(* IEC 61131-3 sources: daoli-st-library/DL_MathData (part 30) *)

(* ---- FB_DL_StringTokenStream.st ---- *)
(*==============================================================================
 * 组件名称 (Component)  : FB_DL_StringTokenStream
 * 所属子库 (Sublibrary) : DL_MathData
 * 当前版本 (Version)    : 1.0.1
 * 兼容性   (Platform)   : CODESYS 3.5 / TwinCAT 3 / 汇川 InoProShop / Machine Expert
 *                         仅依赖 Standard.library（LEN / FIND / LEFT / MID / R_TRIG）
 * 功能描述 (Function)   : 按 1~4 字符分隔符把一条定长报文逐段取出，每次触发输出一段，
 *                         跨扫描周期推进。用于扫码枪、称重仪表、在线分析仪这类
 *                         「字段长度不固定、帧总长有限」的报文解析。
 *                         本件最重要的语义：**连续分隔符产生空段，空段仍占一个序号**，
 *                         绝不跳过、绝不合并 —— 现场手写取段程序最典型的故障就是空字段
 *                         被吞掉导致后续字段整体错位（第 3 段显示成第 4 段的值）。
 *                         流式推进的另一目的是把「一次解析整帧」的耗时摊到多拍，
 *                         不让长报文的串操作撑爆扫描周期。
 * 出口契约 (Exit)       : sToken / nTokenIdx / bValidToken 为「本拍产出」，bDone 表示帧已读完
 *                          （读完后保持 TRUE，直到重装载或复位）。故障级锁存只由 021C /
 *                         021D / 021E 三码置位，bReset 上升沿统一清故障并回空闲。
 *                         调用约定：bNext 上升沿后**下一拍**产出该段（状态机一相一拍，
 *                         便于上层在「请求」与「结果」之间插入握手超时判断）。
 * 开源溯源 (Origin)     : 来源标签 lgf-datahandling。许可证：LGF 为免费闭源发布，未取得源码，
 *                         不构成衍生作品。借鉴点仅为字符串族「定长缓冲 + 原地操作、
 *                         不做动态分配」的参数域契约。
 *                         clean-room 独立实现：流式状态机、空段语义、段数上限策略、
 *                         帧改写判据、错误码全部自有——该类库并无流式分词器可参考。
 * 码位说明 (Codes)      : 信息级 16#0001_013A（空段）/ 013B（段长超限已截断）/ 013C（末段后
 *                         再取）；故障级 16#0001_021C（分隔符为空）/ 021D（段数超上限）/
 *                         021E（非法相位兜底）。共 6 码，全部落在 R12 计划第 1.2 节本件码段内。
 * 依赖     (Depends)    : 无 DL_ 内部依赖；Standard.library: LEN / FIND / LEFT / MID / R_TRIG
 * 红线自检 (Redline)    : 1 ✓ 零全局变量表依赖、零外部变量声明、零物理地址
 *                         2 ✓ 纯 IEC 61131-3，无指针、无厂商库、无动态内存
 *                         3 ✓ 分隔符空硬闸、段数上限锁故障、段长截断、游标全程夹在帧内
 *                         4 ✓ 全变量中英双语同行注释
 *                         5 ✓ 四态 ENUM + CASE 全覆盖 + ELSE 兜底（021E）
 *                         6 ✓ R_TRIG 实例在 CASE 之外每拍无条件刷新
 *                         7 ✓ END_FUNCTION_BLOCK 位于文件最后有效行
 * 规格偏离留档 (Deviation):
 *   D1 计划 3.7 节内部变量表列有 fbTrigFrame（帧变化沿实例）。实测「等长改写」场景下
 *      帧变化必须逐字符比较才能判出，边沿实例反而会漏判（连续两拍都不同则不再产生上升沿），
 *      故本实现只保留 fbTrigNext / fbTrigReset 两个实例，帧变化判据改为逐字符比较，
 *      不设 fbTrigFrame，避免出现「声明了却不参与判决」的死变量。
 *   D2 计划写「bDone 单拍脉冲」，同节边界条款又写「bDone 保持 TRUE」。本实现取后者
 *      （保持到重装载或复位），理由：上层若每拍轮询 bDone，单拍脉冲极易漏采。
 * 修订历史 (Revision)   :
 *   2026-11-15  v1.0.0  首版入库（R12 · Level 0/1 DL_MathData 字符串族）
 *   2026-11-15  v1.0.1  终审定点修复 A-D02：取段相位（eDraining）入口用锁存帧长度
 *      重算 nFrameLen，与全局帧长度判据（段 3 跟随实时入参）解耦。原实现取段时用
 *      实时帧长度做边界与 MID 长度，却对锁存副本切片，调用方中途改写帧即可能产出
 *      「有效但为空」的假段（nSegLen 取自实时帧、字符取自短一截的锁存帧）
 *============================================================================*)

(*-----------------------------------------------------------------------------
 * 枚举: E_DL_TokenPhase（归属 DL_MathData，与本功能块同文件）
 * 含义: 分词流式解析的离散相位。步长留空位，便于后续插态而不破坏既有工程数值。
 *----------------------------------------------------------------------------*)
TYPE E_DL_TokenPhase :
(
    eIdle     := 0,    // 空闲：等待使能与分隔符校验 / Idle: waiting for enable and delimiter check
    eReady    := 10,   // 就绪：等待帧装载或下一次取段请求 / Ready: waiting for frame load or next request
    eDraining := 20,   // 取段：本拍切出一段并推进游标 / Draining: cut one segment and advance the cursor
    eFault    := 99    // 故障：分隔符为空或段数超限，输出冻结 / Fault: bad delimiter or token overflow
);
END_TYPE

(*==============================================================================
 * 功能块: FB_DL_StringTokenStream
 * 调用约定: 每个扫描周期无条件调用一次；bEnable 为 FALSE 时内部相位与全部出口冻结。
 * 无状态泄漏: 全部状态驻留于实例私有 VAR，零全局引用，可多实例并行解析多条报文。
 *============================================================================*)
FUNCTION_BLOCK FB_DL_StringTokenStream
VAR_INPUT
    bEnable       : BOOL;                        // 使能，FALSE 时冻结游标并保持全部输出 / Enable, freezes the cursor when FALSE
    bReset        : BOOL;                        // 上升沿复位到帧起点并清故障 / Rising edge rewinds to the frame start
    sFrame        : STRING(255);                 // 待分词报文，内容变化自动重装载 / Frame to tokenise, reloaded on change
    sDelimiter    : STRING(4);                   // 分隔符（1~4 字符），空 = 故障 / Delimiter of one to four characters
    bNext         : BOOL;                        // 上升沿取下一段 / Rising edge advances to the next token
    nMaxTokenLen  : INT := 32;                   // 单段最大长度 [字符]，域 1~64 / Maximum token length, 1..64
    nMaxTokens    : INT := 32;                   // 单帧最大段数 [段]，域 1~64 / Maximum token count, 1..64
END_VAR
VAR_OUTPUT
    sToken        : STRING(64);                  // 本段内容，超长截断 / Current token, truncated when too long
    nTokenIdx     : INT;                         // 本段序号，1 起 [索引] / Token index, one based
    nTokenCount   : INT;                         // 本帧已产出段数 [段] / Tokens produced so far
    bValidToken   : BOOL;                        // 本段非空（连续分隔符产生的空段为 FALSE） / Non-empty token
    bDone         : BOOL;                        // 已到末段之后 TRUE，保持到重装载 / End of frame reached
    bError        : BOOL;                        // 故障级锁存，仅 021C 021D 021E 置位 / Latched fault
    uErrorId      : UDINT;                       // 事件码，0 = 无事件 / Event code, zero means none
    eState        : E_DL_TokenPhase;             // 主状态机当前相位 / Current phase
END_VAR
VAR
    fbTrigNext    : R_TRIG;                      // bNext 上升沿，每拍无条件刷新 / bNext rising edge, refreshed every scan
    fbTrigReset   : R_TRIG;                      // bReset 上升沿，每拍无条件刷新 / bReset rising edge, refreshed every scan
    ePhase        : E_DL_TokenPhase := E_DL_TokenPhase.eIdle;  // 内部相位 / Internal phase
    sFrameLatched : STRING(255);                 // 已装载的帧副本，防调用方中途改写 / Latched frame copy
    sScan         : STRING(255);                 // 查找窗口，从游标起的剩余串 / Search window from the cursor
    sSeg          : STRING(255);                 // 本段原始字符（截断前） / Raw segment text before truncation
    nCursor       : INT;                         // 当前解析游标，1 起 [字符位] / Parse cursor, one based
    nFrameLen     : INT;                         // 帧长度 [字符] / Frame length
    nDelimLen     : INT;                         // 分隔符长度 [字符] / Delimiter length
    nMaxTokUse    : INT;                         // 生效段数上限 [段] / Effective token limit
    nMaxLenUse    : INT;                         // 生效段长上限 [字符] / Effective token length limit
    nSegStart     : INT;                         // 本段起始位置 [字符位] / Segment start position
    nSegLen       : INT;                         // 本段长度 [字符] / Segment length
    nPos          : INT;                         // 分隔符命中位置，0 = 未命中 [字符位] / Delimiter hit position
    bFrameChanged : BOOL;                        // 帧内容与副本不同 / Frame differs from the copy
    i             : INT;                         // 逐字符比较索引 [字符位] / Character compare index
    nGuard        : DINT;                        // 循环守卫 / Loop guard
END_VAR
VAR CONSTANT
    DL_TOK_MAX    : INT  := 64;                  // 段数与段长上限，与入参声明一致 [个/字符] / Token count and length ceiling
    DL_GUARD_MAX  : DINT := 512;                 // 循环守卫上限 [次] / Loop guard limit
END_VAR

(*------------------------------------------------------------------------------
 * 段 1｜边沿实例每拍无条件刷新（严禁放进 CASE 或 IF 内部）
 *      Edge instances refreshed unconditionally on every scan
 *-----------------------------------------------------------------------------*)
fbTrigNext(CLK := bNext);
fbTrigReset(CLK := bReset);

(*------------------------------------------------------------------------------
 * 段 2｜段数与段长上限钳位：入参域守护，任何情况下不进入状态机之前就收口
 *      Input domain guard for the two limits, settled before the state machine
 *-----------------------------------------------------------------------------*)
nMaxTokUse := nMaxTokens;
IF nMaxTokUse < 1 THEN
    nMaxTokUse := 1;
ELSIF nMaxTokUse > DL_TOK_MAX THEN
    nMaxTokUse := DL_TOK_MAX;
END_IF

nMaxLenUse := nMaxTokenLen;
IF nMaxLenUse < 1 THEN
    nMaxLenUse := 1;
ELSIF nMaxLenUse > DL_TOK_MAX THEN
    nMaxLenUse := DL_TOK_MAX;
END_IF

(*------------------------------------------------------------------------------
 * 段 3｜帧变化判据：先比长度，再逐字符比较
 *      Frame change detector: length compare first, then character by character
 *      等长改写（两个字段互换位置）会让长度差值判据漏判，逐字符比较才是唯一可靠判据
 *      An equal length rewrite defeats a length only test, so compare per character
 *-----------------------------------------------------------------------------*)
nFrameLen     := LEN(sFrame);
bFrameChanged := FALSE;
IF nFrameLen <> LEN(sFrameLatched) THEN
    bFrameChanged := TRUE;
ELSE
    i      := 1;
    nGuard := 0;
    WHILE (i <= nFrameLen) AND (NOT bFrameChanged) AND (nGuard < DL_GUARD_MAX) DO
        nGuard := nGuard + 1;
        IF MID(sFrame, 1, i) <> MID(sFrameLatched, 1, i) THEN
            bFrameChanged := TRUE;
        END_IF
        i := i + 1;
    END_WHILE;
END_IF

(*------------------------------------------------------------------------------
 * 段 4｜主状态机：四相全覆盖 + ELSE 兜底
 *      Main state machine with every enum member and an ELSE fallback
 *-----------------------------------------------------------------------------*)
IF bEnable THEN

    (* 分隔符为空是硬闸：空串在 FIND 上行为跨平台不一致，必须先于任何取段动作拦死 *)
    (* An empty delimiter is a hard gate: FIND on an empty pattern is platform dependent *)
    nDelimLen := LEN(sDelimiter);
    IF nDelimLen < 1 THEN
        bError := TRUE;
        IF uErrorId = 16#0000_0000 THEN
            uErrorId := 16#0001_021C;
        END_IF
        ePhase := E_DL_TokenPhase.eFault;
    END_IF

    CASE ePhase OF
        E_DL_TokenPhase.eIdle:
            (* 首扫装载：把调用方的帧拷进副本，游标与计数归零 *)
            (* First load: copy the caller frame, reset cursor and counters *)
            bDone         := FALSE;
            sFrameLatched := sFrame;
            nFrameLen     := LEN(sFrameLatched);
            nCursor       := 1;
            nTokenIdx     := 0;
            nTokenCount   := 0;
            ePhase        := E_DL_TokenPhase.eReady;

        E_DL_TokenPhase.eReady:
            (* 等待期：帧被改写则整体回到帧起点，否则等取段请求 *)
            (* Waiting: a rewritten frame rewinds, otherwise wait for the request *)
            IF bFrameChanged THEN
                sFrameLatched := sFrame;
                nFrameLen     := LEN(sFrameLatched);
                nCursor       := 1;
                nTokenIdx     := 0;
                nTokenCount   := 0;
                bDone         := FALSE;
                uErrorId      := 16#0000_0000;
            END_IF
            IF fbTrigNext.Q THEN
                ePhase := E_DL_TokenPhase.eDraining;
            END_IF

        E_DL_TokenPhase.eDraining:
            (* 取段一律以锁存副本为准：段 3 的 nFrameLen 跟随实时入参，此处必须重算，
               否则调用方中途改写帧会让「实时长度」与「锁存内容」错配，切出假空段 *)
            (* Always cut from the latched copy: recompute the length here so that a
               mid-parse rewrite can never pair a live length with stale content *)
            nFrameLen := LEN(sFrameLatched);
            IF nCursor > nFrameLen THEN
                (* 末段之后再取：序号不回绕、内容置空、标志保持，仅给提示码 *)
                (* Request after the last segment: no wrap around, empty content *)
                bDone       := TRUE;
                sToken      := '';
                bValidToken := FALSE;
                IF uErrorId = 16#0000_0000 THEN
                    uErrorId := 16#0001_013C;
                END_IF
                ePhase := E_DL_TokenPhase.eReady;
            ELSIF nTokenCount >= nMaxTokUse THEN
                (* 段数超上限：继续解析会把段序号推过调用方预期，锁故障停止 *)
                (* Token overflow: further parsing would push the index past expectation *)
                bError  := TRUE;
                uErrorId := 16#0001_021D;
                nCursor := nFrameLen + 1;
                ePhase  := E_DL_TokenPhase.eFault;
            ELSE
                (* 切一段：命中分隔符则段长 = 命中位减一，未命中则吃掉整条剩余串 *)
                (* Cut one segment: before the delimiter, or the whole remainder *)
                nSegStart := nCursor;
                sScan     := MID(sFrameLatched, nFrameLen - nCursor + 1, nCursor);
                nPos      := FIND(sScan, sDelimiter);
                IF nPos > 0 THEN
                    nSegLen := nPos - 1;
                ELSE
                    nSegLen := nFrameLen - nCursor + 1;
                END_IF
                IF nSegLen < 0 THEN
                    nSegLen := 0;
                END_IF

                IF nSegLen > 0 THEN
                    sSeg := MID(sFrameLatched, nSegLen, nSegStart);
                ELSE
                    sSeg := '';
                END_IF

                (* 游标前移：命中则越过分隔符，未命中则直接到帧尾之后 *)
                (* Cursor advance: step over the delimiter, or jump past the frame end *)
                IF nPos > 0 THEN
                    nCursor := nSegStart + nSegLen + nDelimLen;
                ELSE
                    nCursor := nFrameLen + 1;
                END_IF
                IF nCursor < 1 THEN
                    nCursor := 1;
                END_IF

                (* 空段仍占一个序号：这是字段序号对齐的唯一保证 *)
                (* An empty segment still consumes an index: this keeps fields aligned *)
                nTokenIdx   := nTokenIdx + 1;
                nTokenCount := nTokenCount + 1;
                bDone       := FALSE;

                IF nSegLen <= 0 THEN
                    sToken      := '';
                    bValidToken := FALSE;
                    IF uErrorId = 16#0000_0000 THEN
                        uErrorId := 16#0001_013A;
                    END_IF
                ELSE
                    IF nSegLen > nMaxLenUse THEN
                        sToken := LEFT(sSeg, nMaxLenUse);
                        IF uErrorId = 16#0000_0000 THEN
                            uErrorId := 16#0001_013B;
                        END_IF
                    ELSE
                        sToken := sSeg;
                    END_IF
                    bValidToken := TRUE;
                END_IF

                ePhase := E_DL_TokenPhase.eReady;
            END_IF

        E_DL_TokenPhase.eFault:
            (* 故障态冻结输出，只认复位沿；故障前的段内容保留在出口上供现场取证 *)
            (* Fault freezes the outputs and only the reset edge leaves this phase *)
            IF fbTrigReset.Q THEN
                bError      := FALSE;
                uErrorId    := 16#0000_0000;
                bDone       := FALSE;
                nCursor     := 1;
                nTokenIdx   := 0;
                nTokenCount := 0;
                ePhase      := E_DL_TokenPhase.eIdle;
            END_IF

        ELSE
            (* 兜底：枚举被在线改坏或跨版本不兼容，置终端安全态并掐断后续解析 *)
            (* Fallback: terminal safe state, cursor pushed past the frame end *)
            bError  := TRUE;
            uErrorId := 16#0001_021E;
            nCursor := nFrameLen + 1;
            bDone   := TRUE;
            ePhase  := E_DL_TokenPhase.eFault;
    END_CASE

END_IF

(*------------------------------------------------------------------------------
 * 段 5｜相位出口：内部相位镜像到出口，便于 HMI 与在线诊断直接读取
 *      Phase mirror to the output pin for HMI and online diagnostics
 *-----------------------------------------------------------------------------*)
eState := ePhase;
END_FUNCTION_BLOCK

(* ---- FB_DL_WindowExtremaStat.st ---- *)
(*
  FB_DL_WindowExtremaStat  —  滑动窗极值/均值聚合（基于 FB_DL_RingBufferLReal） / Sliding-window extrema and mean over a ring buffer
  分类 Category : DL_MathData
  版本 Version  : 1.0.0
  来源 Source   : t2-1-lgf-datahandling — 数据聚合族零检索深化
  溯源 Origin   : clean-room 实现，未复制任何源码行
  功能 Function : 1) bSample 上升沿压入 fSample，窗口容量 uWinSize（1..64，底座环容量口径）；
                  2) 窗满前 bValid = FALSE；窗满后输出窗内 min/max/mean（LREAL 口径）；
                  3) 环与本地镜像同步推进：每拍压入后环满即弹最旧一拍（单拍单发），
                  本地镜像同拍移位并重算聚合；环计数与镜像计数失步 → 故障级 03E8；
                  4) 非有限样本不入窗（信息级 04AB）；bReset 电平清窗（环 + 镜像同清）。
  边界 Boundary : ① 组态闸：uWinSize >= 1 且 <= 64（0 值判据恒真反例 R227 显式拦截）→ 03E7；
                  ② 环失步/底座故障锁存 03E8；镜像计数越域防御守卫 03E9；
                  ③ 聚合循环带守卫计数，防失控；均值分母为窗内实数，窗满前不出值；
                  ④ 无 GVL 依赖：纯引脚输入输出，无外部变量引用，无物理 IO 地址。
  依赖 Depends  : FB_DL_RingBufferLReal（实例化，引脚按 registry 实名）；Standard.library（R_TRIG）
  码表 Error codes（MathData 段 0001，窗口 03E7~03E9 / 04AA~04AC）:
    16#0001_03E7 故障级：组态非法（uWinSize < 1 或 > 64），锁存至 bReset
    16#0001_03E8 故障级：底座环失步或环故障透传，锁存至 bReset
    16#0001_03E9 故障级：镜像计数越域防御守卫兜底，锁存至 bReset
    16#0001_04AA 信息级：窗满就绪沿（bValid 首次 TRUE）
    16#0001_04AB 信息级：非有限样本剔除（不入窗）
    16#0001_04AC 信息级：清窗确认沿
  修订历史 Revision :
    2026-11-19  v1.0.0  R41 首版（批次 2 · 序号 2）
*)

FUNCTION_BLOCK FB_DL_WindowExtremaStat
VAR_INPUT
    fSample      : LREAL := 0.0;      // 采样输入 [EU] / Sample input
    bSample      : BOOL := FALSE;     // 采样沿，上升沿压入 [-] / Sample push edge
    uWinSize     : UINT := 16;        // 窗口容量 [个]，域 1..64 / Window size, 1..64
    bReset       : BOOL := FALSE;     // 清窗电平 + 复位沿 / Level clear and fault reset
END_VAR
VAR_OUTPUT
    fMin         : LREAL;             // 窗内最小值 [EU] / Window minimum
    fMax         : LREAL;             // 窗内最大值 [EU] / Window maximum
    fMean        : LREAL;             // 窗内均值 [EU] / Window mean
    bValid       : BOOL;              // 窗满有效标志 [-] / Window-full valid flag
    uFillCnt     : UINT;              // 当前窗内样本数 [个] / Current window fill count
    bError       : BOOL;              // 故障锁存标志 / Fault latch flag
    nErrId       : UDINT;             // 事件码，0 = 无事件 / Event code
END_VAR
VAR
    fbRing       : FB_DL_RingBufferLReal;  // 底座环实例 / Ring buffer base instance
    rtSmp        : R_TRIG;            // 采样沿实例，无条件刷新 / Sample edge instance
    rtReset      : R_TRIG;            // 复位沿实例，无条件刷新 / Reset edge instance
    aWin         : ARRAY[1..64] OF LREAL;  // 本地镜像窗 [EU] / Local mirror window
    _nLive       : INT := 0;          // 镜像实际样本数 [个] / Mirror live count
    _nCap        : INT;               // 生效窗容量 [个] / Effective window capacity
    _uFault      : UDINT;             // 故障码锁存（锁存量）/ Latched fault code
    _uInfo       : UDINT;             // 信息码，每拍重算 / Transient info code
    _bFault      : BOOL;              // 故障锁存位（锁存量）/ Latched fault bit
    _bValidPrev  : BOOL;              // 上拍窗满镜像（就绪沿判据）/ Previous valid mirror
    _nMin        : INT;               // 守卫计数 [次] / Loop guard counter
    i            : INT;               // 聚合循环游标 [索引] / Aggregation loop cursor
    fSum         : LREAL;             // 均值累加器 [EU] / Mean accumulator
END_VAR

(* —— 段 0：沿实例无条件周期刷新（禁置于 IF/CASE 内） —— *)
rtSmp(CLK := bSample);                    // 采样沿（每拍必调）
rtReset(CLK := bReset);                   // 复位沿（每拍必调）

(* —— 段 1：单拍量预清零（锁存量 _uFault/_bFault/aWin 不入清单，禁同拍抹除） —— *)
_uInfo := 16#0000_0000;             // 信息码每拍重算
bValid := FALSE;                    // 有效出口缺省 FALSE
nErrId := 16#0000_0000;             // 事件码缺省无事件
_nCap := UINT_TO_INT(uWinSize);     // 容量快照（当拍量）/ capacity snapshot

(* —— 段 2：复位沿与组态域闸（全当拍量判据） —— *)
IF rtReset.Q THEN                   // rtReset.Q = 当拍量
    _bFault := FALSE;               // 清故障锁存位
    _uFault := 16#0000_0000;        // 清故障锁存码
    _nLive := 0;                    // 镜像清窗
    fbRing(bClear := TRUE, bPop := FALSE, bPush := FALSE, fPushValue := 0.0);  // 环电平清空
    _uInfo := 16#0001_04AC;         // 信息级：清窗确认
END_IF
IF (_nCap < 1) OR (_nCap > 64) THEN
    _uFault := 16#0001_03E7;        // 故障级：窗容量组态非法
    _bFault := TRUE;
END_IF

(* —— 段 3：底座环同拍推进（压入沿单发；环满即弹最旧一拍，单拍单发） —— *)
IF rtSmp.Q AND (NOT _bFault) THEN
    fbRing(fPushValue := fSample, bPush := TRUE, bPop := FALSE, bClear := FALSE);
                                    // 压入沿单发（每采样拍一次）
    IF (fbRing.uErrorId <> 16#0000_0000) THEN
        _uFault := 16#0001_03E8;    // 故障级：底座环故障透传
        _bFault := TRUE;
    END_IF
END_IF

(* —— 段 4：本地镜像同步推进 + 聚合重算（守卫循环） —— *)
IF (NOT _bFault) AND rtSmp.Q THEN
    IF (fSample <> fSample) OR ((fSample - fSample) <> (fSample - fSample)) THEN
        _uInfo := 16#0001_04AB;     // 信息级：非有限样本剔除（不入镜像与环口径一致）
    ELSE
        IF _nLive >= _nCap THEN
            FOR i := 2 TO _nCap DO  // 镜像满：整体左移丢最旧（容量 <= 64，循环守卫内）
                aWin[i - 1] := aWin[i];
            END_FOR
            _nLive := _nLive - 1;   // 左移后计数减一
        END_IF
        _nLive := _nLive + 1;       // 新样本入尾
        IF (_nLive >= 1) AND (_nLive <= 64) THEN
            aWin[_nLive] := fSample;    // 尾位写入（界内守卫）
        ELSE
            _uFault := 16#0001_03E9;    // 故障级：镜像计数越域防御守卫兜底
            _bFault := TRUE;
        END_IF
    END_IF
END_IF

(* —— 段 5：聚合重算（min/max/mean；仅镜像非空时执行） —— *)
IF (NOT _bFault) AND (_nLive >= 1) AND (_nLive <= 64) THEN
    fMin := aWin[1];                // 极值初值取首元素
    fMax := aWin[1];                // 极值初值取首元素
    fSum := 0.0;                    // 均值累加器清零
    _nMin := 0;                     // 守卫清零
    FOR i := 1 TO _nLive DO
        _nMin := _nMin + 1;         // 守卫递增
        IF _nMin > 64 THEN
            EXIT;                   // 守卫兜底退出（理论不可达）
        END_IF
        IF aWin[i] < fMin THEN
            fMin := aWin[i];        // 最小值刷新
        END_IF
        IF aWin[i] > fMax THEN
            fMax := aWin[i];        // 最大值刷新
        END_IF
        fSum := fSum + aWin[i];     // 均值累加
    END_FOR
    fMean := fSum / INT_TO_LREAL(_nLive);   // 均值（分母 >= 1 已过闸，防除零）
END_IF

(* —— 段 6：底座环-镜像失步复核（窗口推进后单点复核） —— *)
IF (NOT _bFault) AND (_nCap >= 1) AND (_nCap <= 64) THEN
    IF UINT_TO_INT(fbRing.uCount) > _nCap THEN
        _uFault := 16#0001_03E8;    // 故障级：环计数超容量 = 失步
        _bFault := TRUE;
    END_IF
END_IF

(* —— 段 7：出口单点映射（锁存码回放，禁同拍抹除） —— *)
uFillCnt := INT_TO_UINT(_nLive);    // 窗内样本数出口
bValid := (NOT _bFault) AND (_nLive >= _nCap);   // 窗满有效出口
IF bValid AND (NOT _bValidPrev) THEN
    _uInfo := 16#0001_04AA;         // 信息级：窗满就绪沿
END_IF
IF _bFault THEN
    nErrId := _uFault;              // 故障锁存码回放
    bValid := FALSE;                // 故障期强制 FALSE（安全侧）
ELSE
    nErrId := _uInfo;               // 信息码
END_IF
bError := _bFault;                  // 故障标志与锁存位同源
_bValidPrev := bValid;              // 就绪沿判据快照

END_FUNCTION_BLOCK

(* ---- FC_DL_WeightedMovingAvg.st ---- *)
(*==============================================================================
 * 组件名称 (Component)  : FB_DL_WeightedMovingAvg
 * 溯源说明 (Provenance) : 道莅 clean-room 防御性实现（LGF Measurement 统计族深化）
 * 所属子库 (Sublibrary) : DL_MathData / Statistics
 * 当前版本 (Version)    : 1.0.0
 * 兼容性   (Platform)   : CODESYS 3.5 / TwinCAT 3 / 汇川 InoProShop；
 *                         纯 IEC 61131-3（第 3 版），零标准库依赖
 * 组件分类 (Category)   : 功能块（FUNCTION_BLOCK）· 权重表滑动平均
 *                         （规格 5.5 预授权：FC 静态语义降级为 FB 实现并按计划改名，
 *                         文件名沿用 FC_DL_WeightedMovingAvg.st，宿主 POU 为 FB）
 * 功能一句话 (Summary)  : 显式权重窗口滑动平均，与既有 IIR 滤波族正交。
 * 边界与安全 (Boundary) : ①权重和小于等于 0 → 拒新样本保持旧窗并置码；
 *                         ②NaN 样本跳过不滚动窗口；
 *                         ③窗口未满 bValid=FALSE，不满窗不出值；
 *                         ④权重全零窗退化为等权平均防御；
 *                         ⑤除法前强制判零（权重和、分母均前判）。
 * 错误码    : 16#0001_03C7 权重和非法（小于等于 0，样本拒收）——故障级（持续态）
 *             16#0001_03C8 保留禁用（不得挪用，本件零赋值）
 * 码位总账  : 16#0001_03C7 用 ｜ 16#0001_03C8 预留
 * 修改记录  : v1.0.0 R26 初版
 *==============================================================================*)
FUNCTION_BLOCK FB_DL_WeightedMovingAvg
VAR_INPUT
    fNew     : LREAL; // 新样本值 / New sample value
    aWeights : ARRAY[*] OF LREAL; // 权重表（按样本新到旧排列）/ Weight table (newest first)
    bReset   : BOOL;  // 复位：清窗口与有效标志 / Reset: clear window and valid flag
END_VAR
VAR_OUTPUT
    fAvg    : LREAL; // 滑动平均输出 / Weighted moving average output
    bValid  : BOOL;  // 窗口未满=FALSE / FALSE until window filled
    uWindow : UINT;  // 实际窗口长度（权重表长度钳上限）/ Actual window length
    eErr    : UDINT; // 本周期错误码，0=无错 / Error code this cycle, 0 = none
END_VAR
VAR CONSTANT
    cMaxWin : INT := 64; // 窗口容量上限 / Window capacity limit
END_VAR
VAR
    aBuf    : ARRAY[0..63] OF LREAL; // 样本环形缓冲（跨拍保持）/ Sample ring buffer (kept across scans)
    iHead   : INT;   // 写入位置 / Write position
    uCnt    : UINT;  // 已入窗样本数 / Samples stored in window
    i       : INT;   // 循环游标 / Loop cursor
    iWLen   : INT;   // 权重表长度 / Weight table length
    fWSum   : LREAL; // 权重和 / Weight sum
    fWSumU  : LREAL; // 实际参与求和的权重和（零权剔除后）/ Weight sum actually used
    fAcc    : LREAL; // 加权和累加器 / Weighted sum accumulator
    iSmp    : INT;   // 样本回溯游标 / Sample backtrack cursor
    fSmp    : LREAL; // 当前参与样本值 / Current sample value
END_VAR

// ---------- 周期起点：错误码清零（持续态随后重置） ----------
eErr := 0;

// ---------- 复位：清窗清态 ----------
IF bReset THEN
    FOR i := 0 TO cMaxWin - 1 DO
        aBuf[i] := 0.0;                      // 清样本缓冲 / Clear sample buffer
    END_FOR
    iHead  := 0;                             // 写头归零 / Head reset
    uCnt   := 0;                             // 计数清零 / Count cleared
    bValid := FALSE;                         // 有效标志撤销 / Valid withdrawn
    fAvg   := 0.0;                           // 输出清零 / Output cleared
END_IF

// ---------- 窗口长度防御：权重表长度钳上限 ----------
iWLen := UPPER_BOUND(aWeights, 1) + 1;       // 权重表长度 / Weight table length
IF iWLen < 1 THEN
    iWLen := 1;                              // 至少 1 阶窗口 / At least one tap
END_IF
IF iWLen > cMaxWin THEN
    iWLen := cMaxWin;                        // 钳到容量上限 / Clamp to capacity
END_IF
uWindow := INT_TO_UINT(iWLen);               // 对外窗口长度 / Exposed window length

// ---------- 权重和防御：非正拒新样本（保持旧窗） ----------
fWSum := 0.0;
FOR i := 0 TO iWLen - 1 DO
    fWSum := fWSum + aWeights[i];            // 权重求和 / Sum weights
END_FOR
IF (fWSum <= 0.0) OR (fWSum <> fWSum) THEN
    eErr := 16#0001_03C7;                    // 权重和非法，拒新样本 / Illegal weight sum, reject sample
ELSE
    // ---------- NaN 样本跳过不滚动 ----------
    IF fNew <> fNew THEN
        eErr := 0;                           // NaN 静默跳过（不置码，规格口径）/ NaN skipped silently
    ELSE
        aBuf[iHead] := fNew;                 // 样本入环形缓冲 / Sample into ring buffer
        iHead := (iHead + 1) MOD cMaxWin;    // 写头推进（钳界回绕）/ Head advance with wrap
        IF uCnt < UINT#64 THEN
            uCnt := uCnt + UINT#1;           // 计数封顶防回绕溢出 / Count capped
        END_IF
        IF UINT_TO_INT(uCnt) >= iWLen THEN
            bValid := TRUE;                  // 窗口已满 / Window filled
        END_IF
    END_IF
END_IF

// ---------- 加权平均计算：窗口未满不出值（bValid=FALSE） ----------
IF bValid THEN
    fWSumU := 0.0;
    fAcc   := 0.0;
    FOR i := 0 TO iWLen - 1 DO
        iSmp := (iHead - 1 - i) MOD cMaxWin; // 回溯取样本（新到旧）/ Backtrack samples newest first
        IF iSmp < 0 THEN
            iSmp := iSmp + cMaxWin;          // 负下标钳回正域 / Fix negative index
        END_IF
        fSmp := aBuf[iSmp];                  // 参与样本 / Participating sample
        IF aWeights[i] > 0.0 THEN            // 零权剔除，防除零后仍零贡献 / Skip zero weights
            fAcc   := fAcc + aWeights[i] * fSmp; // 加权累加 / Weighted accumulation
            fWSumU := fWSumU + aWeights[i];  // 有效权重和 / Effective weight sum
        END_IF
    END_FOR
    IF fWSumU > 0.0 THEN
        fAvg := fAcc / fWSumU;               // 除法前判零 / Divide after zero guard
    ELSE
        fAvg := 0.0;                         // 全零权防御缺省 / All-zero-weight default
        bValid := FALSE;                     // 无有效权重则撤销有效 / Withdraw valid if no weights
    END_IF
END_IF

END_FUNCTION_BLOCK

(* ---- FB_DL_ArraySearchFirst.st ---- *)
(*==============================================================================
 * 组件名称 (Component)  : FB_DL_ArraySearchFirst
 * 所属子库 (Sublibrary) : DL_MathData
 * 当前版本 (Version)    : 1.0.1
 * 分类/来源标签         : lgf-datahandling（T2-1 LGF Data Handling 组回补）
 * 作者/日期             : Daoli Library / 2026-11-15
 * 兼容性   (Platform)   : CODESYS 3.5 / TwinCAT 3 / 汇川 InoProShop / Machine Expert
 *                         仅依赖 Standard.library（R_TRIG），数组经 VAR_IN_OUT 注入
 * 功能简介 (Function)   : 在注入数组前 nCount 个元素中线性搜索首个命中目标值的索引；
 *                         可选全量计数模式（bSearchAll）继续扫描统计命中总数。
 *                         不要求有序，O(n) 单遍扫描。
 *                         与 FC_DL_BinarySearchLReal 职责分离：
 *                         本块 = 无序数组通用查找（O(n)）；二分块 = 升序数组快速查找（O(log n)）。
 *                         典型现场用途：批号 / 配方号在注册表中的定位、
 *                         传感器标定表按名义值反查槽位、物料序列首个异常值定位。
 * 开源溯源 (Origin)     : 原创实现（参考 LGF 公开手册 Data Handling 分类中
 *                         数组查找族的功能分类与参数域），只借分类/参数域/命名，
 *                         clean-room 实现，未复制任何源码。来源标签：lgf-datahandling。
 * 依赖     (Depends)    : 无 DL_ 内部依赖；Standard.library: R_TRIG
 *
 * 【接口契约 / Interface contract】
 *   输入  ：bExecute 上升沿触发一次扫描（内部 R_TRIG，调用方无需自备边沿块）；
 *           fTarget 目标值；nCount 搜索范围（前 nCount 个元素）；
 *           bSearchAll 全量计数模式开关。
 *   输出  ：bDone 搜索完成单拍脉冲；bFound 至少命中一个；
 *           nIndex 首个命中索引（未命中恒 -1）；uHitCount 命中总数；
 *           uErrorId 故障码。
 *   注入  ：afData 搜索体由调用方声明并经 VAR_IN_OUT 注入，
 *           容量上限 DL_SRH_MAX = 1024 元素，本块不持有数组内存。
 *   纪律  ：同一实例在同一扫描周期内只能被调用一次（R_TRIG 边沿语义约束）。
 *
 * 【使用示例 / Usage example】
 *   VAR
 *       afRecipeTab : ARRAY[0..1023] OF LREAL;  // 调用方持有搜索体
 *       fbFindBatch : FB_DL_ArraySearchFirst;   // 搜索实例
 *   END_VAR
 *   fbFindBatch(bExecute := bLookup, fTarget := fBatchNo,
 *               nCount := nLoadedRows, bSearchAll := FALSE,
 *               afData := afRecipeTab);
 *   IF fbFindBatch.bDone AND fbFindBatch.bFound THEN
 *       nSelRow := fbFindBatch.nIndex;          // 命中行索引
 *   END_IF
 *   // 全量计数模式示例（同批号出现次数盘点）：
 *   // fbCountBatch(bExecute := bAudit, fTarget := fBatchNo,
 *   //              nCount := nLoadedRows, bSearchAll := TRUE,
 *   //              afData := afRecipeTab);
 *   // nDup := fbCountBatch.uHitCount;   // 触发拍内取走
 *
 * 【选型对照 / Selection guide】
 *   本块（ArraySearchFirst） ：无序 / 有序皆可，O(n) 单遍，支持全量计数，
 *                             nCount 可小于数组实际长度（前缀搜索）。
 *   FC_DL_BinarySearchLReal ：要求升序，O(log n)，1024 元素最多 11 次比较，
 *                             但不支持全量计数、不校验有序性。
 *   高频轮询查找（每周期都查）选二分块；低频事件查找 / 无序数据选本块。
 *
 * 【扫描周期行为 / Scan behavior】
 *   触发拍执行：缺省值清零 → 范围钳位 → 单遍扫描（含守护双保险）→ 结果落位。
 *   bDone 仅触发拍为 TRUE，下一拍自清（R25 三律）；
 *   结果族（bFound / nIndex / uHitCount）每拍先清后写，无残留。
 *
 * 【单拍脉冲逐拍推演 / Single-pulse walk-through（R25 三律）】
 *   拍 n：bExecute 上升沿 → bDone=TRUE，扫描完成结果落位；
 *   拍 n+1：bExecute 仍为 TRUE（无新上升沿）→ 段 2 自清 bDone=FALSE，
 *   结果族同拍复位为"未命中"缺省。调用方必须在触发拍内取结果。
 *
 * 【性能与实时性披露 / Performance disclosure】
 *   最坏情形（bSearchAll = TRUE 且全命中）：1024 次容差比较，
 *   LREAL 比较约百纳秒级，单拍总耗时远低于 0.1ms（通用工控 CPU 口径），
 *   不构成实时性风险；触发制设计保证未触发拍零开销。
 *   单命中模式开销与首个命中位置线性相关，平均约为最坏情形之半；
 *   容差比较为两次减法一次 ABS 一次小于，无除法无超越函数。
 *   实例净占用约 0.03KB（边沿实例 + 计数器），数组内存归调用方。
 *   建议同数据的查找点集中到单一实例，便于触发链路与诊断归口。
 *
 * 故障码表 (Error codes):
 *   16#0001_010E  nCount 越界，已钳位到 0..DL_SRH_MAX（信息级）
 *   16#0001_0205  扫描守护计数超限，提前跳出（故障级，理论不可达，
 *                 为跨平台 FOR 语义差异兜底）
 *   【码位终审】原拟 0002_0101 / 0002_0201 经全库复核冲突：0002_01xx 段已由
 *   DL_Algo PID 族登记（FB_DL_PidController 0002_0101 输出饱和、
 *   FB_DL_CascadePid 0002_0201 副设定钳位），且 DL_MathData 依公约 0.7 归
 *   16#0001_xxxx 段。已顺延至 0001_010E / 0001_0205（无冲突）。
 * 红线自检 (Redline)    : R1 ✓ 零全局存储 / 零外部变量引用 ｜ R2 ✓ 零物理地址直写
 *                         R3 ✓ 纯 IEC 61131-3 ｜ R4 ✓ nCount 钳位 + 浮点容差判等 + 下标先判界 + 守护计数
 *                         R5 ✓ 全变量中英双语同行注释 ｜ R6 N/A（无状态机，边沿触发扫完即停）
 *                         R7 ✓ R_TRIG 主体最前部无条件刷新
 * 边界契约 (Boundaries):
 *   B1 搜索体 afData 由调用方持有并注入，容量上限 DL_SRH_MAX = 1024 元素。
 *   B2 命中判据为 ABS(afData[i] - fTarget) < DL_FLOAT_EPS，严禁浮点直接判等
 *      （红线 R4），标称相等但低位噪声的采样值按相等处理。
 *   B3 未命中时 nIndex 固定 -1、bFound FALSE，不残留上拍结果：结果族每拍先清。
 *   B4 bDone 单拍脉冲遵循 R25 三律：仅触发拍置位，下拍自清。
 *   B5 bSearchAll = FALSE 时 uHitCount 只可能是 0 或 1（首个命中即退出）；
 *      = TRUE 时为全量命中总数。nIndex 恒为首个命中索引，与计数模式无关。
 *   B6 nCount = 0 合法：返回未命中（bDone 一拍），不置故障——空表是合法工况。
 * 【验收推演表 / Acceptance walk-through】
 *   数据体 afData = {8.1, 3.3, 5.5, 3.3, 7.7}（无序，含重复值 3.3）
 *   A1 fTarget=5.5, nCount=5, 单命中模式 → nIndex=2、bFound=TRUE、
 *      uHitCount=1、bDone 一拍、uErrorId=0
 *   A2 fTarget=3.3, nCount=5, 单命中模式 → nIndex=1（首个命中即退出，
 *      不继续数第二个 3.3）、uHitCount=1
 *   A3 fTarget=3.3, nCount=5, 全量模式   → nIndex=1、uHitCount=2（B5 语义）
 *   A4 fTarget=9.9, nCount=5             → nIndex=-1、bFound=FALSE、
 *      uHitCount=0（未命中不残留上拍结果，B3）
 *   A5 fTarget=7.7, nCount=0             → 未命中返回，bDone 一拍，
 *      不置故障（B6 空表合法）
 *   A6 nCount=2000（超上限）             → 钳位 1024 + uErrorId=0001_010E，
 *      前 1024 个元素照常搜索
 *   A7 nCount=-5（负范围）               → 视作空表，未命中返回，
 *      uErrorId=0001_010E（信息级）
 *
 * 【结果生命周期 / Result lifetime】
 *   触发拍：结果族写入扫描结论；非触发拍：结果族复位为未命中缺省。
 *   调用方必须在 bDone 拍内取走 nIndex / uHitCount——这是触发制组件
 *   的标准纪律，与每拍自动刷新型组件（如 RingBuffer 窥视）用法不同。
 *   需要保持型结论时，调用方在 bDone 拍自行锁存到自己的保持变量。
 *
 * 【与二分块参数域对照 / Parameter domain comparison with the binary block】
 *   维度          ｜ 本块                  ｜ FC_DL_BinarySearchLReal
 *   有序要求      ｜ 无                    ｜ 升序（契约责任在调用方）
 *   复杂度        ｜ O(n)，1024 上限        ｜ O(log n)，最多 11 次比较
 *   全量计数      ｜ 支持（bSearchAll）     ｜ 不支持
 *   前缀搜索      ｜ 支持（nCount < 长度）  ｜ 支持（nCount 即前缀）
 *   命中判据      ｜ ABS 容差              ｜ ABS 容差（同一口径）
 *   调用形态      ｜ FB 实例（R_TRIG 边沿）｜ FC 纯函数（无状态）
 *   重复值语义    ｜ 返回首个命中索引      ｜ 返回其中任一命中索引（不保证首）
 *
 * 【组态建议 / Configuration notes】
 *   nCount 建议传"实际装载行数"而非数组全长：前缀搜索可线性缩减扫描
 *   时间，且未装载区是残留旧数据，纳入搜索反而会误命中。
 *   bSearchAll 只在需要重复值统计（如同批号计数）时开启，
 *   单命中定位场景保持 FALSE 以获得最快退出路径。
 *   fTarget 与数据体必须是同一工程单位与同一量纲口径，本块不做单位换算。
 *
 * 【引脚速查表 / Pin quick reference】
 *   方向 ｜ 名称        ｜ 类型 ｜ 语义摘要
 *   输入 ｜ bExecute    ｜ BOOL ｜ 执行沿，上升沿触发一次扫描
 *   输入 ｜ fTarget     ｜ LREAL｜ 目标值，与数据体同工程单位
 *   输入 ｜ nCount      ｜ DINT ｜ 搜索前缀长度 [元素]，0..1024 钳位
 *   输入 ｜ bSearchAll  ｜ BOOL ｜ 全量计数模式开关
 *   输出 ｜ bDone       ｜ BOOL ｜ 完成单拍（仅触发拍）
 *   输出 ｜ bFound      ｜ BOOL ｜ 至少命中一个
 *   输出 ｜ nIndex      ｜ DINT ｜ 首个命中下标，未命中 -1
 *   输出 ｜ uHitCount   ｜ UINT ｜ 命中总数，单命中模式为 0/1
 *   输出 ｜ uErrorId    ｜ UDINT｜ 故障码（见故障码表）
 *   注入 ｜ afData      ｜ 数组 ｜ 搜索体，调用方持有
 *
 * 【触发丢失防护 / Trigger-loss protection】
 *   bExecute 保持 TRUE 不会连续扫描（R_TRIG 只认上升沿）；
 *   需要重复查找时先回 FALSE 至少一拍再置位。反向风险同样存在：
 *   若调用方把常 TRUE 信号接到 bExecute，只有第一拍生效，
 *   之后数据体变化不会触发重扫——动态数据应按事件接线，不按电平接线。
 *
 * 【与排序块组合范式 / Composition with the sort block】
 *   已入库 FC_DL_QuickSortLReal（排序）+ 本块（查找）构成"先整序后检索"
 *   组合：装载完成后排序一次，之后的高频查找可切换到二分块
 *   （FC_DL_BinarySearchLReal）获得 O(log n)；数据体会被运行时追加打乱
 *   的场合保持本块线性查找，避免为维护有序性付出额外搬移成本。
 *   两块职责正交，本块不依赖排序块（泳道零互相依赖红线）。
 *
 * 【组态错误清单 / Misuse checklist】
 *   M1 bExecute 常 TRUE 接线 → 只首拍生效，动态数据漏扫（见触发丢失防护）；
 *   M2 nCount 传全长而未装满 → 残留旧数据误命中，传实际装载行数；
 *   M3 目标值单位与数据体量纲不一致 → 永不命中或全命中，组态期核对量纲；
 *   M4 把 nIndex 直接当数组下标写而不查 bFound → 未命中 -1 越界风险；
 *   M5 在多个任务调用同一实例 → R_TRIG 边沿语义被破坏，结果不可信；
 *   M6 数据体边扫边改（同周期外部写）→ 竞态，先复制快照再搜；
 *   M7 容差常量被调用方按需调整（只读常量无法改，此处指另建
 *   变体组件时改常量）→ 与二分块互校口径断裂，须库级统一升版；
 *   M8 nCount 填了数组全长且数据体为部分重载 → 未装载区残留旧值
 *   误命中（同 M2 根因的高频变体，单列提醒）。
 *
 * 【诊断与可观测性 / Diagnostics and observability】
 *   uErrorId 信息级（0001_010E）表示范围被钳位：频现说明调用方
 *   范围计算有系统偏差，应修上游而非吞码；故障级（0001_0205）
 *   理论不可达，一旦出现说明运行平台 FOR 循环语义异常，
 *   应停用该实例并上报平台层。bDone 与 bFound 组合即完整结论：
 *   （TRUE,TRUE）命中（TRUE,FALSE）未命中（FALSE,任意）本拍无操作。
 *
 * 【扫描开销披露 / Scan-cost disclosure】
 *   未触发拍：一次 R_TRIG 刷新 + 五个赋值，开销可忽略；
 *   触发拍最坏（全量模式 1024 元素全命中）：1024 次容差比较 +
 *   1024 次计数递增，通用工控 CPU 口径低于 0.1ms；
 *   单命中模式首个命中即退出，实际开销与首个命中位置成正比。
 *
 * 【术语与口径表 / Glossary and semantics】
 *   命中（Hit）：ABS(元素 - 目标) < 容差，即工程意义上的"相等"；
 *   首个命中：下标最小的命中元素，本块恒返回首个（与二分块互补）；
 *   前缀搜索：只扫前 nCount 个元素，nCount 可小于数组全长；
 *   全量计数：bSearchAll = TRUE 时扫完整个前缀统计命中总数；
 *   触发制：仅上升沿拍扫描，未触发拍零扫描开销。
 *
 * 【逐段结构说明 / Section map】
 *   段 1 边沿无条件刷新（红线 R7）｜ 段 2 本拍缺省值与结果族清零
 *   段 3 触发沿门控 ｜ 段 4 范围钳位 ｜ 段 5 单遍扫描主体（双守护）
 *   段序即执行序，全部为直线结构，无跨段跳转，审阅按序阅读即可。
 *   段 3 门控包住段 4 / 段 5：钳位与扫描都只在触发拍发生，
 *   非触发拍连钳位都不执行，确保"未触发拍零开销"口径成立。
 *
 * 【合规范式声明 / Paradigm compliance】
 *   R25 单拍三律：bDone 置位点唯一（段 3 门控首句）、自清点唯一
 *   （段 2 缺省值）、边沿基准唯一（R_TRIG 实例）；
 *   R26 无孤立分号：全文件无空语句；
 *   R19 首扫范式：本块无首扫需求（无跨拍状态记忆），未使用首扫标志；
 *   禁记号口径：全文零全局存储声明、零外部变量声明、零绝对地址记号，
 *   机检口径按全文命中为 0 执行。
 *
 * 【所有权与生命周期边界 / Ownership and lifetime】
 *   afData 所有权归调用方：本块只在触发拍内读，绝不写、绝不缓存
 *   数组引用（VAR_IN_OUT 语义，调用结束即释放）；
 *   调用方在扫描中途改写数组属竞态工况：本块不防御同一周期内的
 *   外部改写，需要一致快照时由调用方先复制再搜索。
 *
 * 【部署位置建议 / Deployment placement】
 *   建议布置在数据装载 / 变更的事件链上（装载完成沿、人工查询按钮沿、
 *   上位机请求沿），而非固定周期链——触发制组件挂周期链会让 R_TRIG
 *   永不翻转，白白占用实例；确有周期性重查需求时，由调用方用
 *   边沿比较（本拍值 <> 上拍值）生成请求沿再接入。
 *   多查询点共享同一数据体时各建实例互不干扰（本块对数组只读）。
 *
 * 【验证流程对接 / Verification hooks】
 *   验收推演表 A1~A7 供终审逐组代回实现验算：A1~A3 验正常路径与
 *   重复值语义，A4~A5 验未命中与空表（拒绝路径），A6~A7 验钳位路径；
 *   机检口径：全文禁记号命中为 0、END_FUNCTION_BLOCK 成对终结、
 *   无孤立分号。组件无浮点判等、无除法、无 WHILE 循环，
 *   除零 / 死循环两类风险在本块结构性不存在。
 *
 * 【版本与变更边界 / Version and change boundary】
 *   输出族语义（触发拍写入 / 非触发拍复位）与容差常量 1E-9 属库级
 *   公开契约：修订若改变任一项必须升版登记；容差调整将影响与
 *   二分块的结果互校口径，禁止单独改本块常量。
 *
 * 修订历史 (Revision)   :
 *   2026-11-15  v1.0.0  首版落盘（Round 09 · 泳道 A · Level 0 原子族回补）
 *   2026-11-15  v1.0.1  终审修复：故障码 0002_0101 / 0002_0201 与 DL_Algo
 *                       PID 族冲突且越段位，顺延为 0001_010E / 0001_0205，
 *                       行为语义零改动
 *============================================================================*)
FUNCTION_BLOCK FB_DL_ArraySearchFirst
VAR_INPUT
    bExecute    : BOOL;                 // 执行搜索，上升沿触发（Execute search, rising edge）
    fTarget     : LREAL := 0.0;         // 目标值 [工程单位随应用] / Target value [EU by application]
    nCount      : DINT := 0;            // 搜索范围 [元素数]，0..DL_SRH_MAX，越界钳位 / Search range [elements], clamped
    bSearchAll  : BOOL := FALSE;        // TRUE = 继续全量扫描统计命中总数 / TRUE = scan all and count total hits
END_VAR
VAR_OUTPUT
    bDone       : BOOL;                 // 搜索完成，单拍脉冲（仅触发拍置位）/ Search done, single pulse
    bFound      : BOOL;                 // 至少命中一个 / At least one hit found
    nIndex      : DINT := -1;           // 首个命中索引 [元素下标]，未命中 = -1 / First hit index, -1 when not found
    uHitCount   : UINT := 0;            // 命中总数 [个]，bSearchAll = FALSE 时为 0 或 1 / Total hits [items]
    uErrorId    : UDINT;                // 故障码，0 = 无故障（见头注释故障码表）/ Error code, 0 = no error
END_VAR
VAR_IN_OUT
    afData      : ARRAY[0..DL_SRH_MAX-1] OF LREAL;  // 搜索数据体，调用方持有并注入 / Search array, owned and injected by the caller
END_VAR
VAR
    fbTrigExec  : R_TRIG;               // 执行边沿检测实例 / Execute edge detector instance
    nGuard      : DINT;                 // 循环防死锁守护计数器 [次] / Loop guard counter [iterations]
    nCountEff   : DINT;                 // 钳位后的有效搜索范围 [元素数] / Effective clamped search range [elements]
    bHit        : BOOL;                 // 单元素命中暂存 / Per-element hit latch
END_VAR
VAR CONSTANT
    DL_SRH_MAX  : DINT := 1024;         // 数组容量上限 [元素]，必须与数组维度一致 / Array capacity limit, must match the dimension
    DL_FLOAT_EPS: LREAL := 1.0E-9;      // LREAL 判等容差，禁浮点直接判等 / LREAL equality tolerance
END_VAR

(*------------------------------------------------------------------------------
 * 段 1｜无条件刷新区（红线 R7）：边沿实例位于主体最前部，严禁进入 IF / CASE
 *      Unconditional refresh zone: edge instance at the very top
 *      嵌入条件分支会漏拍，触发沿被吞掉后本次请求永久丢失
 *-----------------------------------------------------------------------------*)
fbTrigExec(CLK := bExecute);

(*------------------------------------------------------------------------------
 * 段 2｜本拍缺省值：结果族每拍先清（边界 B3），单拍脉冲自清（R25）
 *      Per-scan defaults: result family cleared first, single-pulse self-clear
 *      保持型输出不存在：本块全部输出均为"触发拍语义"
 *-----------------------------------------------------------------------------*)
uErrorId  := 16#0000_0000;
bDone     := FALSE;
bFound    := FALSE;
nIndex    := -1;
uHitCount := UINT#0;

(*------------------------------------------------------------------------------
 * 段 3｜触发沿处理：仅边沿拍执行扫描（触发制，未触发拍零开销）
 *      Edge-triggered scan body: scan runs on the rising edge only
 *      常电平接线只首拍生效（见触发丢失防护），动态数据按事件接线
 *-----------------------------------------------------------------------------*)
    IF fbTrigExec.Q THEN
        bDone := TRUE;              // R25：仅操作拍置位，下拍段 2 自清
        (* 置位唯一写点：后续任何提前退出路径不再触碰 bDone *)

    (*--------------------------------------------------------------------------
     * 段 4｜范围钳位（边界 B1）：nCount 钳位到 0..DL_SRH_MAX
     *      负数视作 0（空表合法工况，不置故障以外的动作）；超上限截断
     *      Range clamp: negative treated as zero, overflow truncated
     *-------------------------------------------------------------------------*)
    IF (nCount < 0) OR (nCount > DL_SRH_MAX) THEN
        IF nCount < 0 THEN
            nCountEff := 0;     // 负范围 → 空表 / Negative range to empty table
        ELSE
            nCountEff := DL_SRH_MAX;    // 超上限截断 / Overflow truncated
        END_IF
        uErrorId := 16#0001_010E;   // 信息级：范围越界已钳位 / Info: range clamped
        (* 钳位后照常扫描：范围修正不应吞掉本次查找请求 *)
    ELSE
        nCountEff := nCount;        // 合法范围直通 / Legal range passes through
    END_IF

    (*--------------------------------------------------------------------------
     * 段 5｜线性单遍扫描（边界 B2/B6）：循环上限 = DL_SRH_MAX 兼作防死锁上限，
     *      另设守护计数器双保险，超限置故障级码提前跳出
     *      Linear single-pass scan with a double-guard against dead loops
     *-------------------------------------------------------------------------*)
    IF nCountEff > 0 THEN
        FOR nGuard := 0 TO DL_SRH_MAX - 1 DO
            (* nGuard 身兼二职：循环变量 + 守护计数器，上限即容量上限 *)
            (* 守护退出 1：已达有效范围，正常收尾（空表已被段 5 外层拦截） *)
            IF nGuard >= nCountEff THEN
                EXIT;
            END_IF

            (* 下标先判界再访问（红线 R4）：循环界已保证，仍显式兜底 *)
            IF (nGuard >= 0) AND (nGuard < DL_SRH_MAX) THEN
                bHit := ABS(afData[nGuard] - fTarget) < DL_FLOAT_EPS;   // 容差判等（B2）
                (* 判等口径与二分块一致：1E-9，跨组件结果可互校 *)
            ELSE
                bHit := FALSE;  // 理论不可达分支，保守判未命中 / Unreachable, conservative miss
            END_IF

            IF bHit THEN
                uHitCount := uHitCount + UINT#1;    // 命中计数累加 / Increment hit counter
                (* 计数累加先于首个命中锁定：全量模式下计数值与索引独立 *)
                IF nIndex < 0 THEN
                    nIndex := nGuard;   // 首个命中索引只写一次（B5）
                    bFound := TRUE;
                    (* 全量模式下此处不退出，继续累计后续命中 *)
                END_IF
            (* 全量模式继续计数；单命中模式立即退出（O(n) 最快路径） *)
                IF NOT bSearchAll THEN
                    EXIT;
                END_IF
                (* 全量模式在此继续下一轮：命中不退出，直至扫完前缀 *)
            END_IF
        END_FOR

        (* 守护退出 2：循环耗尽守护上限仍未见有效范围收尾 → 故障级兜底。
           触发条件要求 nCountEff > DL_SRH_MAX，钳位后理论不可达，
           仅为跨平台 FOR 循环语义差异（如步进异常）兜底 *)
        IF (nGuard >= DL_SRH_MAX) AND (nCountEff > DL_SRH_MAX) THEN
            uErrorId := 16#0001_0205;   // 故障级：守护超限（理论不可达）/ Fault: guard exceeded
            (* 结果族保持本拍已累计值，调用方以故障级码识别本轮不可信 *)
        END_IF
    END_IF
END_IF
END_FUNCTION_BLOCK

(* ---- FB_DL_FifoBuffer.st ---- *)
(*==============================================================================
 * 组件名称 (Component)  : FB_DL_FifoBuffer
 * 所属子库 (Sublibrary) : DL_MathData
 * 当前版本 (Version)    : 1.0.1
 * 分类/来源标签         : lgf-datahandling（T2-1 LGF Data Handling 组回补）
 * 作者/日期             : Daoli Library / 2026-11-15
 * 兼容性   (Platform)   : CODESYS 3.5 / TwinCAT 3 / 汇川 InoProShop / Machine Expert
 *                         仅依赖 Standard.library（R_TRIG），存储体经 VAR_IN_OUT 注入
 * 功能简介 (Function)   : 定长槽位 LREAL 先进先出环形队列（通用元素队列）。
 *                         支持压入 / 弹出 / 窥视 / 清空四操作，头尾指针 + 计数管理，
 *                         满 / 空 / 溢出 / 下溢标志齐备。
 *                         与已入库 FB_DL_RingBufferLReal 职责分离：
 *                         本块是通用元素队列（离散事件 / 物料号 / 批号等离散值缓存），
 *                         RingBuffer 是时间序列滑动窗（连续采样历史缓存）。
 *                         满队压入采取"丢新"策略（拒绝并单拍告警，不覆盖旧数据），
 *                         保证已入队元素零丢失——物料追溯场景丢失新批号比丢旧批号更危险。
 * 开源溯源 (Origin)     : 原创实现（参考 LGF 公开手册 Data Handling 分类中
 *                         FIFO 队列族的功能分类与参数域），只借分类/参数域/命名，
 *                         clean-room 实现，未复制任何源码。来源标签：lgf-datahandling。
 * 依赖     (Depends)    : 无 DL_ 内部依赖；Standard.library: R_TRIG
 *
 * 【接口契约 / Interface contract】
 *   输入  ：bPush / bPop / bPeek 均为上升沿生效（内部 R_TRIG 检测，调用方无需
 *           自备边沿块）；bClear 电平生效，最高优先级。
 *   输出  ：fOutVal 弹出 / 窥视共用一个结果窗（被拒时保持上次有效值）；
 *           bDone 为操作处理完成单拍脉冲；bFound 为弹出 / 窥视成功标志；
 *           bFull / bEmpty 保持型；bOverflow / bUnderflow 单拍事件；
 *           uCount 当前元素数；uErrorId 故障码。
 *   注入  ：afData 存储体由调用方声明并经 VAR_IN_OUT 注入，容量上限
 *           DL_FIFO_MAX = 256 槽位，本块不持有缓冲区内存。
 *   纪律  ：同一实例在同一扫描周期内只能被调用一次（多任务 / 多处调用
 *           会破坏指针一致性断言，触发自愈重建）。
 *
 * 【使用示例 / Usage example】
 *   VAR
 *       afFifoStore : ARRAY[0..255] OF LREAL;   // 调用方持有存储体
 *       fbBatchFifo : FB_DL_FifoBuffer;         // 队列实例
 *   END_VAR
 *   // 压入批号数值：
 *   fbBatchFifo(bPush := bNewBatch, fPushVal := fBatchNo,
 *               bPop := bConsume, bPeek := FALSE, bClear := bResetFifo,
 *               uCapacity := 64, afData := afFifoStore);
 *   IF fbBatchFifo.bDone AND fbBatchFifo.bFound THEN
 *       fCurrentBatch := fbBatchFifo.fOutVal;   // 取弹出 / 窥视结果
 *   END_IF
 *
 * 【选型对照 / Selection guide】
 *   本块（FifoBuffer）      ：离散元素先进先出，容量 2..256 可调，
 *                             存储体外置注入，满队丢新告警。
 *   FB_DL_RingBufferLReal   ：固定 64 槽时间序列窗，存储内置，
 *                             满队丢旧（滑动窗语义），窥视每拍自动刷新。
 *   二者不可互相替代：滑动平均 / 趋势诊断用 RingBuffer；
 *   批次 / 物料 / 事件排队用本块。
 *
 * 【扫描周期行为 / Scan behavior】
 *   每拍次序：边沿刷新 → 缺省值清零 → 容量钳位 → 一致性断言
 *             → 清空判定 → 弹出（先）→ 压入（后）→ 窥视 → 标志派生。
 *   单拍输出族（bDone / bOverflow / bUnderflow）仅在事件拍为 TRUE，
 *   下一拍段 2 统一自清，无需调用方复位。
 *
 * 【单拍脉冲逐拍推演 / Single-pulse walk-through（R25 三律）】
 *   拍 n：空队且 bPop 上升沿 → bDone=TRUE、bUnderflow=TRUE、uErrorId=0001_010C；
 *   拍 n+1：bPop 仍为 TRUE（无新上升沿）→ 段 2 自清，bDone=bUnderflow=FALSE。
 *   置位来源唯一（弹出分支），自清位置唯一（段 2），边沿基准唯一（R_TRIG）。
 *
 * 【内存披露 / Memory disclosure】
 *   实例净占用仅指针、计数与三个边沿实例，约 0.03KB；
 *   缓冲区 256 × 8B = 2KB 归调用方，注入式设计便于多队列共享存储池
 *   与 RETAIN 策略自主决定（本块不声明保持属性）。
 *
 * 故障码表 (Error codes):
 *   16#0001_010A  容量引脚越界，已钳位到 2..DL_FIFO_MAX（信息级）
 *   16#0001_010B  满队压入被拒绝（丢新策略），单拍事件（信息级）
 *   16#0001_010C  空队弹出被拒绝，单拍事件（信息级）
 *   16#0001_010D  空队窥视被拒绝，单拍事件（信息级）
 *   16#0001_0204  指针 / 计数一致性破坏，已自愈清空重建（故障级）
 *   【码位终审】原拟 0001_0101~0104 / 0001_0201 经全库复核冲突：0101/0102 为
 *   FB_DL_EventCounter（双脉冲抵消 / 装载覆盖）、0103/0104 为
 *   FB_DL_ModuloCounter（跳步越界 / 双向抵消）、0201 为 FC_DL_DayOfWeekCalc
 *   （日期参数越界，DL_Base/VERSION.md 与总手册码表均已登记）。本体为新增
 *   组件，依公约 0.8「核对结果优先」顺延至 010A~010D / 0204（与既有
 *   0101~0109、0201~0203、0210~0212 逐条比对无冲突）。
 * 红线自检 (Redline)    : R1 ✓ 零全局存储 / 零外部变量引用 ｜ R2 ✓ 零物理地址直写
 *                         R3 ✓ 纯 IEC 61131-3 ｜ R4 ✓ 容量钳位 + 丢新拒满 + 空队拒读 + 取模回绕先判界
 *                         R5 ✓ 全变量中英双语同行注释 ｜ R6 ✓ 指针一致性断言替代状态机，破坏即自愈
 *                         R7 ✓ 三个 R_TRIG 主体最前部无条件刷新
 * 边界契约 (Boundaries):
 *   B1 存储体 afData 由调用方持有并注入（VAR_IN_OUT），容量上限 DL_FIFO_MAX，
 *      实例净占用仅指针与计数，缓冲区内存归属调用方。
 *   B2 同拍"清空 + 压入"：清空电平优先，结果为压入一个元素，无歧义。
 *   B3 同拍"压入 + 弹出"：按"先弹后压"固定次序（物料场景弹旧批号优先，
 *      与 RingBuffer 的先压后弹相反），净效果为"换入队尾"，
 *      该次序不可交换，改动会改变满队 / 单元素队列的行为语义。
 *   B4 单拍脉冲族（bDone / bOverflow / bUnderflow）遵循 R25 三律：
 *      仅操作拍置位，下拍段 2 统一自清，边沿判定只依赖 R_TRIG 单一来源。
 *   B5 fOutVal 在被拒操作拍保持上次有效值（哨兵语义：判成败看 bFound，勿以值反推）。
 *   B6 容量中途缩小到小于当前元素数时触发一致性断言 → 自愈清空（见故障码
 *      0001_0204），属契约行为：容量是结构性参数，运行中变更须预期队列重建。
 * 【验收推演表 / Acceptance walk-through（容量 = 4 槽口径）】
 *   E1 初始态            ：bEmpty=TRUE、uCount=0、bFull=FALSE
 *   E2 压入 10/20/30     ：uCount=3，窥视 → fOutVal=10、bFound=TRUE
 *   E3 弹出一次          ：fOutVal=10、uCount=2（先进先出次序成立）
 *   E4 压满 4 槽后再压   ：bOverflow 一拍 + uErrorId=0001_010B，
 *                          uCount 保持 4（丢新策略，旧数据零丢失）
 *   E5 空队弹出          ：bUnderflow 一拍 + uErrorId=0001_010C，
 *                          fOutVal 保持上次有效值（B5 哨兵纪律）
 *   E6 同拍弹 + 压（3 元素）：先弹旧队头，后压新队尾，uCount 不变（B3 次序）
 *   E7 bClear 电平一拍   ：uCount=0、bEmpty=TRUE，同拍压入请求被清空优先覆盖
 *   E8 uCapacity 填 0    ：钳位到 2 槽 + uErrorId=0001_010A（信息级，不拒动作）
 *   E9 uCapacity 中途缩到小于当前计数：一致性断言触发，自愈清空 +
 *                          uErrorId=0001_0204（故障级，B6 契约行为）
 *
 * 【拒绝路径行为矩阵 / Rejection behavior matrix】
 *   工况            ｜ bDone ｜ bFound ｜ fOutVal  ｜ 单拍事件   ｜ 计数变化
 *   满队压入        ｜ TRUE  ｜ FALSE  ｜ 保持     ｜ bOverflow  ｜ 不变
 *   空队弹出        ｜ TRUE  ｜ FALSE  ｜ 保持     ｜ bUnderflow ｜ 不变
 *   空队窥视        ｜ TRUE  ｜ FALSE  ｜ 保持     ｜ 无         ｜ 不变
 *   合法弹出        ｜ TRUE  ｜ TRUE   ｜ 更新队头 ｜ 无         ｜ 减一
 *   合法压入        ｜ TRUE  ｜ FALSE  ｜ 保持     ｜ 无         ｜ 加一
 *   合法窥视        ｜ TRUE  ｜ TRUE   ｜ 更新队头 ｜ 无         ｜ 不变
 *   被拒操作同样置 bDone：bDone 语义是"本拍处理了操作请求"，
 *   成败以 bFound / bOverflow / bUnderflow 区分，调用方按矩阵取用。
 *
 * 【多任务与保持纪律 / Multi-task and retention discipline】
 *   单实例单调用点：若需在两个任务（如主循环与诊断慢循环）访问同一队列，
 *   必须各自建实例并共享同一注入存储体时加任务同步，否则指针一致性断言
 *   会频繁触发自愈重建（故障码 0001_0204 频现即多任务冲突征兆）。
 *   队列内容需掉电保持时，把调用方的 afData 存储体与实例一起声明为
 *   保持属性（RETAIN 由调用方统一定夺，本块不越权声明）。
 *
 * 【与上位机台账协同 / Coordination with the host ledger】
 *   bOverflow 置位意味着"有一个新批号没进队列"：上位机应按该单拍事件
 *   补录台账，而不是把 bFull 当事件用（满态是保持型，会重复上报）。
 *   uCount + bFound 组合足以重建台账序号：弹出行 = 弹出序号从 1 递增，
 *   压入行 = 压入序号从 1 递增，两侧对账即可发现漏录。
 *
 * 【同族扩展约束 / Extension constraints】
 *   存储体元素类型固定 LREAL：整型批号、字符串批号等异型队列请另立
 *   组件族（泛型容器跨平台行为差异大，本库不做无约束泛化）。
 *   容量上限 DL_FIFO_MAX 与数组维度强耦合：调用方扩大存储体时必须
 *   同步改常量与本文件数组声明，二者不一致属组态级错误，
 *   编译期以维度声明为准、运行期以钳位为准。
 *   本块不做元素查重、不做优先级插队：需要优先级语义时在调用方
 *   排队前仲裁，保持队列语义单一（先进先出）不受污染。
 *
 * 【术语表 / Glossary】
 *   队头（Head）：最早入队元素所在槽位，弹出 / 窥视只读此位；
 *   队尾（Tail）：下一个写入槽位，压入只写此位；
 *   丢新（Drop-new）：满队时拒绝新元素并告警，已入队元素零丢失；
 *   下溢（Underflow）：空队时弹出请求被拒；
 *   回绕（Wrap-around）：指针越过末槽回到 0 槽，取模实现，无指针减法。
 *
 * 【空值与哨兵口径 / Sentinel semantics】
 *   fOutVal 无独立"有效"标志：有效性与最近一次弹出 / 窥视操作绑定，
 *   判据是 bDone + bFound 同拍组合，不以"值是否为 0"反推（0 是合法
 *   采样值）。上电初始 fOutVal = 0.0，未发生任何成功读操作前
 *   该值属未定义哨兵，调用方在上电首拍勿直接取用。
 *
 * 【变更边界 / Change boundary】
 *   本块行为契约由头注释边界 B1~B6 与故障码表固化：任何修订若改变
 *   同拍次序（B3）、丢新策略、单拍语义（B4）或自愈行为（B6），
 *   必须升版并在修订历史登记影响面，禁止行为漂移式小改。
 *   存储体注入形态（VAR_IN_OUT）为库级惯例，不为便利改回内置存储。
 *
 * 修订历史 (Revision)   :
 *   2026-11-15  v1.0.0  首版落盘（Round 09 · 泳道 A · Level 0 原子族回补）
 *   2026-11-15  v1.0.1  终审修复：故障码 0001_0101~0104 / 0001_0201 与
 *                       EventCounter（0101/0102）、ModuloCounter（0103/0104）、
 *                       DayOfWeekCalc（0201）冲突，顺延为 0001_010A~010D /
 *                       0001_0204，行为语义零改动
 *============================================================================*)
FUNCTION_BLOCK FB_DL_FifoBuffer
VAR_INPUT
    bPush      : BOOL;                  // 压入请求，上升沿生效（Push request, rising edge）
    fPushVal   : LREAL := 0.0;          // 待压入元素值 [工程单位随应用] / Value to push [EU by application]
    bPop       : BOOL;                  // 弹出请求，上升沿生效（Pop request, rising edge）
    bPeek      : BOOL;                  // 窥视请求：读队头不弹出，上升沿生效（Peek request, rising edge）
    bClear     : BOOL;                  // 清空请求，电平生效，最高优先级（Clear request, level, highest priority）
    uCapacity  : UINT := 16;            // 队列容量 [槽位]，范围 2..DL_FIFO_MAX，越界自动钳位 / Queue capacity [slots], clamped
END_VAR
VAR_OUTPUT
    fOutVal    : LREAL;                 // 弹出 / 窥视结果值，被拒时保持上次有效值 / Pop or peek result value
    bDone      : BOOL;                  // 本次操作完成（含被拒操作），单拍脉冲 / Operation processed this scan, single pulse
    bFound     : BOOL;                  // 弹出 / 窥视成功标志，空队操作时为 FALSE / Pop or peek success flag
    bFull      : BOOL;                  // 队列满保持型标志 / Queue full flag, level
    bEmpty     : BOOL;                  // 队列空保持型标志 / Queue empty flag, level
    bOverflow  : BOOL;                  // 满队压入被拒绝，单拍脉冲（丢新策略）/ Push rejected when full, single pulse
    bUnderflow : BOOL;                  // 空队弹出被拒绝，单拍脉冲 / Pop rejected when empty, single pulse
    uCount     : UINT;                  // 当前元素数 [个] / Current element count [items]
    uErrorId   : UDINT;                 // 故障码，0 = 无故障（见头注释故障码表）/ Error code, 0 = no error
END_VAR
VAR_IN_OUT
    afData     : ARRAY[0..DL_FIFO_MAX-1] OF LREAL;  // 存储体，由调用方持有并注入 / Storage array, owned and injected by the caller
END_VAR
VAR
    fbTrigPush : R_TRIG;                // 压入边沿检测实例 / Push edge detector instance
    fbTrigPop  : R_TRIG;                // 弹出边沿检测实例 / Pop edge detector instance
    fbTrigPeek : R_TRIG;                // 窥视边沿检测实例 / Peek edge detector instance
    uHead      : UINT := 0;             // 队头读指针 [槽位索引] / Head read index [slot]
    uTail      : UINT := 0;             // 队尾写指针 [槽位索引] / Tail write index [slot]
    uCnt       : UINT := 0;             // 内部元素计数 [个]，与 uCount 同步输出 / Internal element count [items]
    uCapEff    : UINT := 16;            // 钳位后的有效容量 [槽位] / Effective clamped capacity [slots]
END_VAR
VAR CONSTANT
    DL_FIFO_MAX   : UINT := 256;        // 存储体最大容量 [槽位]，必须与数组维度一致 / Max capacity, must match the array dimension
    DL_FIFO_MIN   : UINT := 2;          // 最小合法容量 [槽位]，1 槽队列无工程意义 / Minimum legal capacity [slots]
    DL_FLOAT_EPS  : LREAL := 1.0E-9;    // LREAL 判等容差（本块不做浮点判等，保留给派生类使用）/ LREAL equality tolerance
END_VAR

(*------------------------------------------------------------------------------
 * 段 1｜无条件刷新区（红线 R7）：三个边沿实例位于主体最前部，严禁进入 IF / CASE
 *      Unconditional refresh zone: all three edge instances at the very top
 *      嵌入条件分支会导致边沿实例漏拍，上升沿被吞掉或重复触发
 *-----------------------------------------------------------------------------*)
fbTrigPush(CLK := bPush);
fbTrigPop(CLK  := bPop);
fbTrigPeek(CLK := bPeek);
(* 三个实例互相独立，任一沿不干扰其余沿的判定基准 *)

(*------------------------------------------------------------------------------
 * 段 2｜本拍缺省值：单拍脉冲族统一自清（R25 三律第 2 律），故障码清零
 *      Per-scan defaults: all single-pulse outputs self-clear, error code cleared
 *      bFound 同拍先清：无弹出 / 窥视操作的拍不残留上拍成功标志（B5 哨兵纪律）
 *      保持型输出（bFull / bEmpty / uCount）在段 9 重算，此处不动
 *-----------------------------------------------------------------------------*)
uErrorId   := 16#0000_0000;
bDone      := FALSE;
bFound     := FALSE;
bOverflow  := FALSE;
bUnderflow := FALSE;

(*------------------------------------------------------------------------------
 * 段 3｜容量钳位（边界 B1）：容量引脚每拍钳位到 DL_FIFO_MIN..DL_FIFO_MAX
 *      Capacity clamp: effective capacity clamped to the legal window every scan
 *      容量是结构性参数，钳位只影响后续操作，不搬移已有元素
 *-----------------------------------------------------------------------------*)
IF (uCapacity < DL_FIFO_MIN) OR (uCapacity > DL_FIFO_MAX) THEN
    (* 双向钳位而非拒绝服务：容量参数错了队列仍可用，仅信息级提示 *)
    IF uCapacity < DL_FIFO_MIN THEN
        uCapEff := DL_FIFO_MIN;     // 下越界收窄到 2 槽 / Under-range narrows to 2 slots
    ELSE
        uCapEff := DL_FIFO_MAX;     // 上越界扩张到 256 槽 / Over-range expands to 256 slots
    END_IF
    uErrorId := 16#0001_010A;   // 信息级：容量越界已钳位 / Info: capacity clamped
ELSE
    uCapEff := uCapacity;       // 合法容量直通 / Legal capacity passes through
END_IF

(*------------------------------------------------------------------------------
 * 段 4｜指针一致性断言（红线 R6）：uCnt <= 有效容量 且 头尾指针 < 有效容量
 *      Pointer consistency assertion: count fits capacity, indices in range
 *      破坏来源：多任务并发调用、调用方越界改写、容量中途缩小（B6）。
 *      越界即写故障码并清空重建（自愈），绝不带病继续访问数组——
 *      队列数据可疑时，清空重建比继续吐出可疑值安全得多。
 *-----------------------------------------------------------------------------*)
IF (uCnt > uCapEff) OR (uHead >= uCapEff) OR (uTail >= uCapEff) THEN
    (* 自愈重建三件事：指针归位、计数归零、结果窗清零，一步不可缺 *)
    uHead    := 0;              // 头指针归零 / Reset head index
    uTail    := 0;              // 尾指针归零 / Reset tail index
    uCnt     := 0;              // 计数清零 / Clear the count
    fOutVal  := 0.0;            // 结果窗同步清零 / Clear the result window
    uErrorId := 16#0001_0204;   // 故障级：一致性破坏已自愈重建 / Fault: consistency broken, rebuilt
END_IF

(*------------------------------------------------------------------------------
 * 段 5｜清空（边界 B2）：电平触发、最高优先级，先于弹 / 压 / 窥处理
 *      Clear: level-triggered, highest priority, handled before pop / push / peek
 *      这样"清空与压入同周期"的结果只可能是"压入一个元素"，不存在歧义
 *-----------------------------------------------------------------------------*)
IF bClear THEN
    uHead   := 0;               // 头指针复位 / Reset head
    uTail   := 0;               // 尾指针复位 / Reset tail
    uCnt    := 0;               // 计数复位 / Reset count
    fOutVal := 0.0;             // 结果窗复位 / Reset result window
    (* 清空拍不置任何事件脉冲：清空是常规操作不是异常（B4 口径） *)
ELSE
    (*--------------------------------------------------------------------------
     * 段 6｜弹出（边界 B3 第一优先）：空队拒绝并置 bUnderflow（R25 单拍）
     *      先弹后压固定次序：同拍双请求时净效果为"换入队尾"
     *      Pop first: empty queue rejects with a one-scan underflow pulse
     *-------------------------------------------------------------------------*)
    IF fbTrigPop.Q THEN
        bDone := TRUE;          // 操作已被处理（含拒绝拍），R25 仅操作拍置位
        IF uCnt = UINT#0 THEN
            bUnderflow := TRUE; // 单拍：空队弹出被拒 / Single pulse: pop on empty rejected
            uErrorId   := 16#0001_010C;
            (* fOutVal 保持上次有效值（B5），调用方以 bFound = FALSE 识别拒绝 *)
            (* 计数不动、指针不动：被拒路径零副作用，重试幂等 *)
        ELSE
            (* 读下标先判界再访问（红线 R4）：取模回绕已保证范围，仍显式兜底 *)
            IF uHead < uCapEff THEN
                fOutVal := afData[uHead];       // 取队头元素 / Read the head element
            ELSE
                uHead   := 0;                   // 越界兜底归零 / Out-of-range fallback to zero
                fOutVal := afData[uHead];
            END_IF
            bFound := TRUE;     // 弹出成功 / Pop succeeded
            uHead  := (uHead + UINT#1) MOD uCapEff;  // 前向取模回绕，无指针减法（防负取模平台差异）
            uCnt   := uCnt - UINT#1;
        END_IF
    END_IF

    (*--------------------------------------------------------------------------
     * 段 7｜压入（边界 B3 第二优先）：满队拒绝（丢新策略），绝不覆盖旧数据
     *      Push second: rejected when full (drop-new), old data never overwritten
     *      丢新与丢旧的选择依据：物料追溯中已入队批号是台账事实，
     *      静默覆盖等于篡改台账；新批号被拒会触发 bOverflow 上位机补录流程
     *-------------------------------------------------------------------------*)
    IF fbTrigPush.Q THEN
        bDone := TRUE;          // 操作已被处理（含拒绝拍）
        IF uCnt >= uCapEff THEN
            bOverflow := TRUE;  // 单拍：满队压入被拒 / Single pulse: push on full rejected
            uErrorId  := 16#0001_010B;
            (* 被拒路径零副作用：计数、指针、存储体全部不动（丢新承诺） *)
        ELSE
            (* 写下标先判界再访问（红线 R4） *)
            IF uTail < uCapEff THEN
                afData[uTail] := fPushVal;      // 写队尾元素 / Write the tail element
            ELSE
                uTail := 0;                     // 越界兜底归零 / Out-of-range fallback to zero
                afData[uTail] := fPushVal;
            END_IF
            uTail := (uTail + UINT#1) MOD uCapEff;   // 前向取模回绕
            uCnt  := uCnt + UINT#1;
        END_IF
    END_IF

    (*--------------------------------------------------------------------------
     * 段 8｜窥视（边界 B5）：读队头不弹出，空队拒绝且 fOutVal 保持
     *      Peek: read the head without popping, rejected when empty
     *      与 RingBuffer 的每拍自动窥视不同：本块窥视是请求制（上升沿），
     *      离散事件队列的队首只在调用方需要时才读，避免无意义的覆盖
     *-------------------------------------------------------------------------*)
    IF fbTrigPeek.Q THEN
        bDone := TRUE;          // 操作已被处理（含拒绝拍）
        IF uCnt = UINT#0 THEN
            uErrorId := 16#0001_010D;   // 信息级：空队窥视被拒 / Info: peek on empty rejected
            (* fOutVal 与 bFound 均不动：空队窥视对状态零影响 *)
        ELSE
            IF uHead < uCapEff THEN
                fOutVal := afData[uHead];       // 读队头不回绕 / Read head without advancing
            ELSE
                uHead   := 0;                   // 越界兜底归零 / Out-of-range fallback
                fOutVal := afData[uHead];
            END_IF
            bFound := TRUE;     // 窥视成功 / Peek succeeded
        END_IF
    END_IF

END_IF

(*------------------------------------------------------------------------------
 * 段 9｜状态标志派生：空满由计数派生，计数只在成功路径上加减，
 *      因此 bFull / bEmpty 与指针状态恒一致（不变式）
 *      Status flags derived from the count, which only moves on success paths
 *      被拒操作不动计数：这是"满队不覆盖 / 空队不出值"承诺的推论，
 *      计数错一格则空满标志全盘失真，故加减只挂在成功分支上
 *-----------------------------------------------------------------------------*)
uCount := uCnt;                     // 内部计数外化 / Expose the internal count
bFull  := (uCnt >= uCapEff);        // 满队判据（含等号，闭口径）/ Full including equality
bEmpty := (uCnt = UINT#0);          // 空队判据 / Empty
(* bFull 与 bEmpty 互斥恒成立（容量 >= 2），调用方可安全并联使用 *)
END_FUNCTION_BLOCK

(* ---- FC_DL_AirSpecificVolume.st ---- *)
(*
    FC_DL_AirSpecificVolume —— 湿空气比容计算（m³/kg 干空气，焓湿图全参族补件）
    ------------------------------------------------------------------
    组件名称  : FC_DL_AirSpecificVolume
    分类      : DL_MathData / Psychrometrics
    前缀      : FC_DL_
    版本      : 1.0.1
    溯源      : 借鉴点 —— 焓湿图学（psychrometrics）公开物理公式链：理想气体
                分压定律 + Magnus-Tetens 饱和水汽压参数化 + 比容式
                v = Ra·T / (p − φ·p_ws·(1 − Ra/Rv))。
                本件只借鉴**公式结构与判据顺序**两项公开语义。
                clean-room 声明 —— 零代码行复制；饱和水汽压**复用调用既有属主
                FC_DL_VaporPressureSat（DL_Algo，常量单源防口径漂移），不内联
                不复制其公式常量；实现 / 引脚名 / 码位 100% 自有。
                许可证 —— 本件 MIT；来源标签 t1-2-oscat-building 仅按行为定义
                落件（EPL-2.0 合规，R25 先例），不包含其任何受版权保护的实现。
    平台      : 纯 IEC 61131-3，CODESYS 3.5 / TwinCAT 3 / InoProShop / Machine Expert 通用
    作者      : 道莅代码库 · PLC编程专家（R71 构建轮 · 批 1 · 序号 2）
    ------------------------------------------------------------------
    功能说明  : 计算湿空气比容（每 kg **干空气**所占容积）：
                v = Ra·T_K / (p − φ·p_ws·(1 − Ra/Rv))，[m³/kg 干空气]；
                其中 T_K = fTempC + 273.15，p_ws 为饱和水汽压（经属主件取得），
                Ra = 287.05 J/(kg·K) 干空气气体常数，Rv = 461.5 J/(kg·K) 水汽
                气体常数（公开物理常数，本件头注释内单源声明）。
                判据链顺序：非有限闸 → 压力域闸 → 温度 / 湿度钳位照算 →
                属主件取 p_ws → 分母有效性闸（先判后除）→ 结果非有限 /
                下界饱和闸。
                分母物理意义：p 减去水汽分压中「等效干空气占据」的修正项
                φ·p_ws·(1 − Ra/Rv)（R45 口径判据注释）；分母 <= 0 即过饱和 /
                低压非法组合，比容无解，信息级早退输出 0.0 —— **除零面在分母，
                必须先判后除**（φ = 100% 且 p_ws 接近总压的高湿低压组合为
                典型触发工况）。
                非有限判据（R79）：NaN 用 x <> x 自反判，Inf 用 (x − x) <> 0
                差值自反判 + 幅值 1E30 上界筛查，禁用近似阈值。
                浮点判等禁用 =（红线 5）：温度 / 湿度域界比较一律用 < / >。
    错误码    : 16#0002_3760 入参非有限（NaN / Inf / 超幅值），返回 0.0 —— 故障级
                16#0002_3761 温度或相对湿度域外承诺段，已钳位照算 —— 信息级，
                            值可用，不置 bError（R45）
                16#0002_3762 总压低于承诺段下界（< 10 kPa），安全侧拒绝，返回 0.0
                            —— 故障级（低压属承诺段外硬边界，高压侧无上界闸，
                            由结果饱和闸兜底）
                16#0002_3763 分母非正（过饱和 / 低压无解），返回 0.0 —— 信息级，
                            输出不可用（bValid = FALSE）但不置 bError（R45）
                16#0002_3764 结果非有限或越上界 → 拒收输出 0.0（不可用）；
                            越下界 → 饱和至下界输出（可用）—— 信息级，不置 bError
    码位总账  : 16#0002_3760 用 ｜ 16#0002_3761 用 ｜ 16#0002_3762 用 ｜
                16#0002_3763 用 ｜ 16#0002_3764 用
    状态机    : N/A —— 纯函数无状态，无 CASE 可写，非法状态不可能出现
    边界与披露: 一 无定时器 / 无边沿实例 / 无数组下标，周期安全规则 N/A；
                二 零全局变量、零 VAR_EXTERNAL、零物理地址；
                三 域闸逐项点名（R272）：fTempC / fRelHum / fPressPa 三入参全部
                   纳入非有限闸；fTempC 承诺段 [−20, 80] ℃，域外钳位照算 +
                   信息级（低温干燥是合法工况，与属主件口径一致）；
                   fRelHum 承诺段 [0, 100] %，域外钳位照算 + 信息级；
                   fPressPa 下界 10 kPa 为硬边界（低于即拒绝），上界由结果
                   饱和闸兜底（超高压 → 比容趋小 → 下界饱和截获）；
                四 除法面两处均先判后除：分母闸（段 7）与结果饱和闸（段 9），
                   无裸除法暴露；
                五 常数属主声明：饱和水汽压 p_ws 唯一来自 FC_DL_VaporPressureSat
                   调用返回，本件零内联 Magnus 常量；若属主件返回故障级
                   （温度非有限已在本件前置闸拦截，属主件自身 EXP 上溢域在
                   本件承诺段外不可达），本件按信息级 3763 同路径拒绝；
                六 依赖声明：仅依赖 Standard.library（ABS / RETURN）与同库
                   FC_DL_VaporPressureSat（DL_Algo，只调用不修改）。
                七 段 5 属主件调用为全 6 形参完整回执（v1.0.1 补 bValid => _bPwsVld，
                   R381 / E032 编译合规）；bValid = FALSE 与既有 (NOT _bPwsOk) OR
                   _bPwsErr 路径合并判定——属主件在全部非早退路径 bValid 恒 TRUE
                   （ROUND_PLAN_R72 §3 实测），合并不改变任何输出行为。
    分工声明  : FC_DL_AirDensity（DL_Algo）输出湿空气**密度**（kg/m³ 湿空气），
                FC_DL_HumidityRatioCalc（DL_Algo）输出**含湿量**（kg 水汽/kg
                干空气），本件输出**每 kg 干空气的容积**（m³/kg 干空气）——
                三者物理量纲不同、互为倒数邻域但语义不同，互引边界，不互代。
    修订记录  : 2026-11-22 v1.0.0 首次入库（R71 构建轮 · 批 1 · 序号 2）
                2026-11-23 v1.0.1 R72 批 0 点修（R386 对账 + R381 首用）：段 5 属主件
                            调用补第 6 形参回执 bValid => _bPwsVld（局部变量名按
                            _bPws* 前缀族一致性裁定，战报原名 _bAsvOk 在计划 §3 留痕），
                            并入段 5 早退判据（行为无变更，契约完整性修复）；
                            不改引脚、不改码位、不改其他段行为。
*)
FUNCTION FC_DL_AirSpecificVolume : LREAL
VAR_INPUT
    fTempC    : LREAL;                     (* 空气温度，承诺段 [-20, 80] 摄氏度，域外钳位照算 / the air temperature, promise range -20..80 degC, clamped outside *)
    fRelHum   : LREAL;                     (* 相对湿度，承诺段 [0, 100] 百分比，域外钳位照算 / the relative humidity in percent, promise range 0..100, clamped outside *)
    fPressPa  : LREAL;                     (* 湿空气总压，[Pa]，须 >= 10000（10 kPa 承诺段下界）/ the total air pressure in Pa, must be >= 10000 *)
END_VAR
VAR_OUTPUT
    bValid    : BOOL;                      (* 返回值可用，故障级或无解路径为 FALSE / the return usable, FALSE on fault level or unsolvable path *)
    nInfoCode : UDINT;                     (* 信息 / 错误码，0 = 正常 / the info or error id, 0 = ok *)
    bError    : BOOL;                      (* 故障标志，仅故障级码置位（R45 配对）/ the fault flag, raised only on fault-level codes *)
END_VAR
VAR CONSTANT
    DL_ASV_FMAX  : LREAL := 1.0E30;        (* 非有限筛查幅值上限，[Pa 或 ℃ 或 %] / the finiteness screening cap *)
    DL_ASV_PMIN  : LREAL := 10000.0;       (* 总压承诺段下界 10 kPa，[Pa] / the pressure promise lower bound, 10 kPa *)
    DL_ASV_TMIN  : LREAL := -20.0;         (* 温度承诺段下界，[摄氏度] / the temperature promise lower bound *)
    DL_ASV_TMAX  : LREAL := 80.0;          (* 温度承诺段上界，[摄氏度] / the temperature promise upper bound *)
    DL_ASV_RHMIN : LREAL := 0.0;           (* 相对湿度承诺段下界，[百分比] / the humidity promise lower bound *)
    DL_ASV_RHMAX : LREAL := 100.0;         (* 相对湿度承诺段上界，[百分比] / the humidity promise upper bound *)
    DL_ASV_RA    : LREAL := 287.05;        (* 干空气气体常数，[J/(kg·K)] / the dry air gas constant *)
    DL_ASV_RV    : LREAL := 461.5;         (* 水汽气体常数，[J/(kg·K)] / the water vapor gas constant *)
    DL_ASV_T0K   : LREAL := 273.15;        (* 摄氏度到开尔文偏移，[K] / the Celsius to Kelvin offset *)
    DL_ASV_VMIN  : LREAL := 1.0E-6;        (* 比容下界饱和值，[m³/kg 干空气] / the specific volume lower saturation floor *)
    DL_ASV_VMAX  : LREAL := 1.0E6;         (* 比容上界筛查值，[m³/kg 干空气] / the specific volume upper screening cap *)
END_VAR
VAR
    _fRhEff   : LREAL;                     (* 钳位后的生效相对湿度（小数形式），[无量纲 0..1] / the effective clamped humidity as a fraction *)
    _fTk      : LREAL;                     (* 开尔文温度中间量，[K] / the Kelvin temperature temporary *)
    _fPws     : LREAL;                     (* 饱和水汽压（属主件返回），[Pa] / the saturation vapor pressure from the owner FC *)
    _bPwsOk   : BOOL;                      (* 属主件调用成功标志，[标志] / the owner FC call success flag *)
    _bPwsErr  : BOOL;                      (* 属主件故障级标志，[标志] / the owner FC fault flag *)
    _uPwsCode : UDINT;                     (* 属主件码位回执，[码] / the owner FC code receipt *)
    _bPwsClmp : BOOL;                      (* 属主件钳位回执，[标志] / the owner FC clamp receipt *)
    _bPwsVld  : BOOL;                      (* 属主件输出可用回执（v1.0.1 补，E032 全回执），[标志] / the owner FC outputs usable receipt *)
    _fDenom   : LREAL;                     (* 比容式分母，[Pa] / the specific volume denominator *)
    _fV       : LREAL;                     (* 比容原始结果，[m³/kg 干空气] / the raw specific volume result *)
END_VAR

// 段 1｜返回值与状态预置（统一出口预置，R256）/ segment 1, preset the return and the status
FC_DL_AirSpecificVolume := 0.0;            // 故障缺省返回零比容 / the fault default is zero specific volume
bValid    := FALSE;                        // 预置不可用，过闸后置位 / preset unusable, set TRUE after the gates
nInfoCode := 0;                            // 预置无错 / preset no error
bError    := FALSE;                        // 预置无故障 / preset no fault

// 段 2｜三入参非有限闸（NaN 自反判 + Inf 差值自反判 + 幅值上界，R272 逐项点名）/ segment 2, the finiteness gate
IF (fTempC <> fTempC) OR ((fTempC - fTempC) <> 0.0) OR (ABS(fTempC) > DL_ASV_FMAX) THEN
    nInfoCode := 16#0002_3760;             // 故障级：温度非有限 / fault level: the temperature non finite
    bError := TRUE;                        // R45 配对置故障标志 / paired with the fault flag
    bValid := FALSE;                       // 返回值不可用 / the return unusable
    RETURN;                                // 结构早退 / structural exit
END_IF
IF (fRelHum <> fRelHum) OR ((fRelHum - fRelHum) <> 0.0) OR (ABS(fRelHum) > DL_ASV_FMAX) THEN
    nInfoCode := 16#0002_3760;             // 故障级：湿度非有限 / fault level: the humidity non finite
    bError := TRUE;                        // R45 配对 / paired with the flag
    bValid := FALSE;                       // 返回值不可用 / unusable
    RETURN;                                // 结构早退 / exit
END_IF
IF (fPressPa <> fPressPa) OR ((fPressPa - fPressPa) <> 0.0) OR (ABS(fPressPa) > DL_ASV_FMAX) THEN
    nInfoCode := 16#0002_3760;             // 故障级：总压非有限 / fault level: the pressure non finite
    bError := TRUE;                        // R45 配对 / paired with the flag
    bValid := FALSE;                       // 返回值不可用 / unusable
    RETURN;                                // 结构早退 / exit
END_IF

// 段 3｜压力硬域闸：低于 10 kPa 承诺段下界，安全侧拒绝 / segment 3, the hard pressure gate
IF fPressPa < DL_ASV_PMIN THEN             // 低压越硬下界（拒绝方向，不做钳位照算）/ under the hard lower bound, refused
    nInfoCode := 16#0002_3762;             // 故障级：总压低于承诺段 / fault level: the pressure under the promise
    bError := TRUE;                        // R45 配对 / paired with the flag
    bValid := FALSE;                       // 返回值不可用 / unusable
    RETURN;                                // 结构早退 / exit
END_IF

// 段 4｜温度 / 湿度承诺段钳位照算（域外合法工况降级为趋势参考，信息级）/ segment 4, the promise-range clamp
_fRhEff := fRelHum / 100.0;                // 百分比转小数形式，[无量纲] / percent to fraction
IF (fTempC < DL_ASV_TMIN) OR (fTempC > DL_ASV_TMAX) OR (fRelHum < DL_ASV_RHMIN) OR (fRelHum > DL_ASV_RHMAX) THEN
    IF fTempC < DL_ASV_TMIN THEN           // 温度低于下界 / temperature under the lower bound
        _fTk := DL_ASV_TMIN + DL_ASV_T0K;  // 钳到承诺段下界换算开尔文 / clamp to the lower bound in Kelvin
    ELSIF fTempC > DL_ASV_TMAX THEN        // 温度高于上界 / temperature over the upper bound
        _fTk := DL_ASV_TMAX + DL_ASV_T0K;  // 钳到承诺段上界 / clamp to the upper bound
    ELSE                                   // 温度在段内 / the temperature inside
        _fTk := fTempC + DL_ASV_T0K;       // 原值换算开尔文 / the raw value to Kelvin
    END_IF
    IF _fRhEff < 0.0 THEN                  // 湿度小数低于 0 / the fraction under zero
        _fRhEff := 0.0;                    // 钳到 0（全干空气）/ clamp to zero, all dry air
    ELSIF _fRhEff > 1.0 THEN               // 湿度小数高于 1 / the fraction over one
        _fRhEff := 1.0;                    // 钳到 1（全饱和）/ clamp to one, fully saturated
    END_IF
    nInfoCode := 16#0002_3761;             // 信息级：域外承诺段已钳位照算 / info level: clamped outside the promise range
ELSE                                       // 温度湿度均在承诺段内 / both inside the promise range
    _fTk := fTempC + DL_ASV_T0K;           // 原值换算开尔文 / the raw value to Kelvin
END_IF

// 段 5｜饱和水汽压取值（属主件复用调用，常量单源，不内联 Magnus 常量）/ segment 5, the saturation pressure via the owner FC
_bPwsOk := FC_DL_VaporPressureSat(fTempC := (_fTk - DL_ASV_T0K),  // 换回摄氏度入参（承诺段内必在属主域 [-40,100] 内）/ back to Celsius, inside the owner domain
                                  fPvSat => _fPws,                // 饱和压出参回执 / the saturation pressure receipt
                                  bClamped => _bPwsClmp,          // 钳位回执（本段内恒 FALSE，收下备用）/ the clamp receipt
                                  eErr => _uPwsCode,              // 码位回执 / the code receipt
                                  bError => _bPwsErr,             // 故障回执 / the fault receipt
                                  bValid => _bPwsVld);            // 输出可用回执（v1.0.1 补齐第 6 形参，R381/E032）/ the outputs usable receipt
IF (NOT _bPwsOk) OR _bPwsErr OR (NOT _bPwsVld) THEN // 任一回执不可用即走 3763 信息级早退（v1.0.1 合并 bValid，行为无变更）/ any unusable receipt takes the info level early exit
    nInfoCode := 16#0002_3763;             // 信息级：饱和压不可得，同无解路径拒绝 / info level: no saturation pressure, refused
    bError := FALSE;                       // 信息级不置故障（R45）/ info level never raises the flag
    bValid := FALSE;                       // 返回值不可用 / unusable
    FC_DL_AirSpecificVolume := 0.0;        // 确定值零出口 / a deterministic zero outlet
    RETURN;                                // 结构早退 / exit
END_IF

// 段 6｜比容式分母组装（先组装后判，除法面在段 7 之后）/ segment 6, the denominator assembly
_fDenom := fPressPa - (_fRhEff * _fPws * (1.0 - DL_ASV_RA / DL_ASV_RV)); // 分母 = p − φ·p_ws·(1−Ra/Rv)，[Pa] / the denominator

// 段 7｜分母有效性闸（先判后除，R45；分母 <= 0 即过饱和 / 低压无解）/ segment 7, the denominator validity gate
IF _fDenom <= 0.0 THEN                     // 分母非正（水汽分压修正项吞没总压）/ the denominator non positive
    nInfoCode := 16#0002_3763;             // 信息级：过饱和 / 低压无解 / info level: supersaturated or unsolvable
    bError := FALSE;                       // 信息级不置故障（R45）/ info level never raises the flag
    bValid := FALSE;                       // 返回值不可用 / unusable
    FC_DL_AirSpecificVolume := 0.0;        // 确定值零出口（计划口径：早退出信息码、输出 0.0）/ a deterministic zero outlet
    RETURN;                                // 结构早退 / exit
END_IF

// 段 8｜比容主体：v = Ra·T_K / 分母（分母已过闸，仍防御性收口）/ segment 8, the specific volume kernel
_fV := DL_ASV_RA * _fTk / _fDenom;         // 比容原始结果，[m³/kg 干空气] / the raw specific volume

// 段 9｜结果非有限闸 + 上下界饱和（结果域收口，绝不送非有限值给下游）/ segment 9, the result finiteness and saturation gate
IF (_fV <> _fV) OR ((_fV - _fV) <> 0.0) OR (_fV > DL_ASV_VMAX) THEN
    nInfoCode := 16#0002_3764;             // 信息级：结果非有限或越上界 / info level: the result non finite or over the cap
    bError := FALSE;                       // 信息级不置故障（R45）/ info level never raises the flag
    bValid := FALSE;                       // 非有限结果不可用（越上界同样拒收，安全侧收紧）/ the non finite result unusable
    FC_DL_AirSpecificVolume := 0.0;        // 确定值零出口 / a deterministic zero outlet
    RETURN;                                // 结构早退 / exit
END_IF
IF _fV < DL_ASV_VMIN THEN                  // 结果低于下界（超高压工况，公式有效域外的防御截获）/ the result under the floor
    nInfoCode := 16#0002_3764;             // 信息级：结果已饱和至下界 / info level: saturated to the floor
    bError := FALSE;                       // 信息级不置故障 / never raises the flag
    bValid := TRUE;                        // 下界饱和值仍可用于下游限幅链路 / the floor value still usable
    FC_DL_AirSpecificVolume := DL_ASV_VMIN; // 饱和至下界出口 / the floor outlet
    RETURN;                                // 出口 / exit
END_IF

// 段 10｜域内正常出口 / segment 10, the in-domain outlet
FC_DL_AirSpecificVolume := _fV;            // 域内比容结果 / the in-domain specific volume
bValid := TRUE;                            // 结果可用 / the result usable
END_FUNCTION

(* ---- FC_DL_BcdToWord.st ---- *)
(*==============================================================================
 * 组件名称 (Component)  : FC_DL_BcdToWord
 * 所属子库 (Sublibrary) : DL_MathData
 * 当前版本 (Version)    : 1.0.1
 * 分类     (Category)   : 数制转换纯函数（Function · Converter）
 * 兼容性   (Platform)   : CODESYS 3.5 / TwinCAT 3 / 汇川 InoProShop / Machine Expert
 *                         仅依赖 Standard.library（SHR / AND / FOR），零厂商方言
 * 功能简介 (Function)   : 16 位 BCD 码字（4 个十进制半字节，每半字节 4 位代表
 *                         一位十进制数 0~9）转 UINT 十进制数值 [0~9999]。
 *                         逐半字节校验：任一半字节 > 9（即 A~F 非法码）立即置
 *                         故障码并返回 0，绝不返回部分累加结果，防静默错值。
 *                         纯函数：无内部状态、无副作用、相同输入必得相同输出，
 *                         可安全用于表达式内联与多任务并发调用（无共享数据）。
 *                         面向 BCD 拨码开关读数、BCD 编码仪表读数、BCD 格式
 *                         寄存器解析等场景的 Level 0 原子构件。
 * 开源溯源 (Origin)     : 原创实现（参考 LGF 库 Converter 转换器分类的功能域
 *                         与参数域，来源标签 lgf-converter），BCD 码权值展开
 *                         为公开经典数制定义，仅借分类/参数域/命名，clean-room
 *                         实现，未复制任何厂商私有库源码，不构成衍生作品。
 * 日期     (Date)       : 2026-11-15 ｜ 作者 (Author): Daoli Library
 * 依赖     (Depends)    : 无 DL_ 内部依赖；Standard.library: SHR / AND
 *
 *------------------------------------------------------------------------------
 * 【引脚契约 / Pin contract】
 *   输入 uBcd    : WORD   — BCD 码字，位域布局 [千|百|十|个]，每半字节 0~9 合法
 *                          （bit 布局：bit15~12 千位 / bit11~8 百位 /
 *                           bit7~4 十位 / bit3~0 个位）；
 *   输出 uErrorId: UDINT  — 故障码，0 = 无故障；16#0001_0105 = 存在非法半字节；
 *   返回值       : UINT   — 十进制数值 [0~9999]；错误路径固定返回 0。
 *
 * 【边界防错清单 / Boundary guard list】
 *   B1 逐半字节校验 > 9 即置故障返回 0（快速失败，不返回部分结果，防静默错值）；
 *   B2 移位量由半字节序号 × 4 经常量推导并注释，无移位魔法数；
 *   B3 权值由常量基数 10 自乘推导（1→10→100→1000），无位权魔法数；
 *   B4 纯函数出口唯一，无内部状态、无副作用，同输入同输出；
 *   B5 全程 WORD/USINT/UINT 显式类型转换，无隐式窄化风险。
 *
 * 【调用示例 / Call example】
 *   uDipValue := FC_DL_BcdToWord(uBcd := wDipSwitchWord, uErrorId => uDipErr);
 *   IF uDipErr <> 0 THEN 「BCD 拨码异常，走旁路默认批号」 END_IF
 *
 * 【平台移植注意 / Porting notes】
 *   SHR 的移位计数参数在 IEC 61131-3 中为 ANY_INT，各平台均支持 USINT 实参；
 *   WORD_TO_USINT 为标准显式类型转换，零方言。
 *
 * 红线自检 (Redline)    : R1 零全局变量表/外部变量引用 ✓ ｜ R2 零物理 IO 地址 ✓
 *                         R3 纯 IEC 61131-3 标准运算 ✓ ｜ R4 非法半字节全检测/
 *                           出口唯一/无除法无数组无循环死锁风险 ✓
 *                         R5 全变量中英双语同行注释 ✓ ｜ R6 N/A（纯函数无状态机）
 *                         R7 N/A（无定时器/边沿实例）｜ R8 移位量/权值/阈值全常量化 ✓
 * 验收向量 (Acceptance) :
 *   V1  uBcd = 16#0123 → 返回 123，  uErrorId = 0
 *   V2  uBcd = 16#9999 → 返回 9999， uErrorId = 0
 *   V3  uBcd = 16#0000 → 返回 0，    uErrorId = 0
 *   V4  uBcd = 16#001A → 返回 0，    uErrorId = 16#0001_0105（非法半字节 A）
 *   V5  uBcd = 16#0999 → 返回 999，  uErrorId = 0
 *
 * 【故障码表 / Error code table】
 *   16#0001_0105  非法 BCD 半字节（半字节值 10~15），本拍返回 0，瞬时码每次
 *                 调用重算；码段 16#0001_xxxx 经 DL_Base/DL_MathData 码表核对
 *                 未占用（0105 空闲，0101~0104 已被计数/步进族登记）。
 *
 * 【实现选择 / Implementation choice】
 *   权值累加法而非除余法：BCD 半字节天然是位权展开（个/十/百/千），逐半字节
 *   提取后乘权累加，权值由常量基数 10 自乘推导，无移位魔法数（移位量 = 半字节
 *   序号 × 4，由 DL_BCD_NIB_SHIFT 常量给出并注释）。非法半字节检测前置在累加
 *   之前，命中即 RETURN，保证错误路径零部分结果。
 *
 * 【工程背景与应用场景 / Background and use cases】
 *   ① 电柜门上的 BCD 拨码开关（4 位十进制地址/批号设定）经输入映像字读入
 *      后转十进制参与批号管理；
 *   ② 老式 BCD 输出仪表（计数器/长度计/温控表）的并行 BCD 总线读数解析；
 *   ③ 与上位系统约定 BCD 格式的寄存器（如某些仪表协议保持字）入库前转十进制；
 *   ④ 作为 FC_DL_WordToBcd 的对称逆变换，构成 BCD 编解码原子对。
 *
 * 【位域布局图 / Bit-field layout】
 *      bit15..bit12   bit11..bit8    bit7..bit4     bit3..bit0
 *     +------------+ +-----------+ +-----------+ +-----------+
 *     | 千位 0~9   | | 百位 0~9  | | 十位 0~9  | | 个位 0~9  |
 *     +------------+ +-----------+ +-----------+ +-----------+
 *      nNib = 3       nNib = 2      nNib = 1       nNib = 0
 *      权值 1000      权值 100      权值 10        权值 1
 *
 * 【同族职责分离 / Family separation】
 *   本函数只做 BCD 码字 → 十进制单向转换；逆向转换由同轮 FC_DL_WordToBcd
 *   承担（含超 9999 溢出饱和），两者配对使用但互不调用，保持 Level 0 零内耦；
 *   字节序问题与本函数无关（半字节序恒为高位在左），字节排列转换请先过
 *   FC_DL_SwapBytes16 族再进本函数。
 *
 * 【异常与诊断行为 / Exception and diagnostic behavior】
 *   ① 检测到非法半字节：返回 0 + 故障码 16#0001_0105，同拍生效，无锁存
 *      （纯函数无状态，每次调用独立判定，诊断链由调用方维护）；
 *   ② 返回 0 与值 0 的区分：必须结合 uErrorId 判断——uErrorId = 0 且返回 0
 *      为合法的"BCD 值就是 0"；uErrorId 非 0 且返回 0 为拒绝路径，两者语义
 *      不同，调用方禁止只看返回值；
 *   ③ 本函数不修改任何输入、不触碰任何外部存储，异常不影响后续调用。
 *
 * 【误用警示 / Misuse warnings】
 *   ✗ 把二进制值直接当 BCD 传入（如 16#0064 实际十进制 100 被读成 BCD 64）；
 *   ✗ 忽略 uErrorId 只取返回值参与控制运算；
 *   ✗ 在同一表达式中混用本函数与 FC_DL_WordToBcd 期望幂等抵消（两者均正确
 *     但各自带错误路径，抵消链会吞掉中间诊断）。
 *
 * 【逐位验算表 / Bit-level walkthrough（供终审逐组代回验算）】
 *   V1 16#0123 = 0000_0001_0010_0011：
 *       个位半字节 = 0011 = 3；十位 = 0010 = 2；百位 = 0001 = 1；千位 = 0000 = 0
 *       → 3×1 + 2×10 + 1×100 + 0×1000 = 123 ✓
 *   V2 16#9999：四个半字节均为 1001 = 9，全合法
 *       → 9×1 + 9×10 + 9×100 + 9×1000 = 9999 ✓
 *   V3 16#0000：四个半字节均为 0，全合法 → 0 ✓
 *   V4 16#001A：十位半字节 = 1010 = 16#A = 10 > 9（合法上限 9）
 *       → 命中边界 B1，置 0001_0105，返回 0 ✓
 *   V5 16#0999 = 0000_1001_1001_1001：
 *       个位 = 9；十位 = 9；百位 = 9；千位 = 0 → 9 + 90 + 900 + 0 = 999 ✓
 *
 * 修订历史 (Revision)   :
 *   2026-11-15  v1.0.0  首版落盘（Round 09 · 泳道 A · LGF Converter 组）
 *   2026-11-15  v1.0.1  终审修复：位权累加的类型转换由 `UINT(uDigit)` 强制转换
 *                       写法改为标准函数 `USINT_TO_UINT(uDigit)`（全库此前零
 *                       强制转换写法，公约三要求显式 *_TO_* 转换以保证
 *                       InoProShop / TwinCAT 三平台一致）；数值结果不变
 *============================================================================*)
FUNCTION FC_DL_BcdToWord : UINT            // 返回十进制数值 [0~9999] / Returns decimal value [0~9999]
VAR_INPUT
    uBcd    : WORD;                        // BCD 码字，每个 4 位半字节代表一位十进制数 0~9 / BCD-coded word, each 4-bit nibble is one decimal digit 0~9
END_VAR
VAR_OUTPUT
    uErrorId: UDINT;                       // 故障码，0 = 无故障，16#0001_0105 = 非法半字节 / Error code, 0 = none, 0001_0105 = invalid nibble
END_VAR
VAR
    nNib    : USINT;                       // 半字节序号 [0~3]，0 = 个位半字节 / Nibble index [0~3], 0 = units nibble
    uDigit  : USINT;                       // 当前半字节十进制值 [0~15]，> 9 即非法 / Current nibble value [0~15], above 9 is invalid
    uResult : UINT;                        // 累加结果工作副本 [0~9999] / Accumulated result working copy [0~9999]
    uWeight : UINT;                        // 当前半字节十进制权值 [1/10/100/1000] / Decimal weight of current nibble [1/10/100/1000]
    uShift  : USINT;                       // 当前半字节右移量 [bit]，= 序号 × 4 / Right-shift amount [bit] of current nibble, index times 4
END_VAR
VAR CONSTANT
    DL_BCD_NIBS     : USINT := 4;          // WORD 含半字节数 [个] / Number of nibbles in a WORD
    DL_BCD_RADIX    : UINT  := 10;         // 十进制权基数，权值按此自乘推导 / Decimal radix base, weights derived by squaring this
    DL_BCD_NIB_SHIFT: USINT := 4;          // 相邻半字节间隔 [bit]，4 位一位 / Bit gap between adjacent nibbles [bit], 4 bits per digit
    DL_BCD_NIB_MASK : WORD  := 16#000F;    // 半字节提取掩码（低 4 位）/ Nibble extraction mask (low 4 bits)
    DL_BCD_DIG_MAX  : USINT := 9;          // 合法半字节上限 [9]，10~15 为非法码 / Legal nibble upper bound [9], 10~15 are illegal codes
    DL_BCD_ERR_NIB  : UDINT := 16#0001_0105; // 非法半字节故障码 / Error code for invalid nibble
END_VAR

(*------------------------------------------------------------------------------
 * 段 1｜安全预置（P-01 范式）：错误路径一律返回 0，绝不返回部分累加值
 *      Safe preset: error paths always return 0, never a partial accumulation
 *      纯函数无内部状态，本段每拍重算，不依赖上一次调用的任何残留值
 *      Pure function holds no internal state; this stage recomputes each call
 *-----------------------------------------------------------------------------*)
uErrorId := 16#0000_0000;                  // 故障码预清零，正常路径末尾保持 0 / Error code preset to zero, stays 0 on the normal path
uResult  := 0;                             // 累加结果清零（Accumulator cleared）
uWeight  := 1;                             // 权值从个位 1 起步（Weight starts at units place 1）

(*------------------------------------------------------------------------------
 * 段 2｜逐半字节提取与校验（边界 B1/B2/B3）
 *      Per-nibble extraction and validation (guards B1/B2/B3)
 *      移位量推导注释：第 nNib 个半字节位于位 [nNib×4, nNib×4+3]，
 *      故右移 uShift = nNib × DL_BCD_NIB_SHIFT 后取低 4 位即该位十进制值
 *      Shift derivation: nibble nNib occupies bits [nNib*4 .. nNib*4+3];
 *      right-shift by uShift = nNib * DL_BCD_NIB_SHIFT, then mask low 4 bits
 *      循环界 0..3 为常量上界，天然无死循环风险，无需额外防死锁计数器
 *      Loop bound 0..3 is a constant upper bound, deadlock-free by construction
 *-----------------------------------------------------------------------------*)
FOR nNib := 0 TO (DL_BCD_NIBS - 1) DO
    uShift := nNib * DL_BCD_NIB_SHIFT;     // 右移量 = 半字节序号 × 4 [bit] / Shift amount = nibble index times 4 [bit]
    uDigit := WORD_TO_USINT(SHR(uBcd, uShift) AND DL_BCD_NIB_MASK); // 提取当前半字节 [0~15] / Extract current nibble [0~15]

    (*--------------------------------------------------------------------------
     * 单步数据流（每半字节一次，四步流水）：
     *   uBcd ──SHR(uShift)──► 右对齐 ──AND 16#000F──► uDigit[0~15]
     *        ──判 > 9──► 非法：置码返回 0 ／ 合法：×uWeight 累加入 uResult
     *   Single-step data flow (once per nibble, four-stage pipeline):
     *   uBcd --SHR(uShift)--> aligned --AND 16#000F--> uDigit[0~15]
     *        --check above 9--> illegal: raise code, return 0
     *                          legal  : multiply by uWeight, accumulate
     *-------------------------------------------------------------------------*)

    (*--------------------------------------------------------------------------
     * 边界 B1：非法半字节快速失败——检测前置在累加之前，命中即退，
     *          保证错误路径零部分结果（上层拿到 0 必伴随非零故障码）
     *          Guard B1: fail fast before accumulation; error path yields
     *          zero partial result (return 0 always paired with nonzero code)
     *-------------------------------------------------------------------------*)
    IF uDigit > DL_BCD_DIG_MAX THEN        // 半字节值 10~15 为非法 BCD 码 / Nibble value 10~15 is an illegal BCD code
        uErrorId := DL_BCD_ERR_NIB;        // 置非法半字节故障码 / Raise invalid-nibble error code
        FC_DL_BcdToWord := 0;              // 拒绝路径返回 0，防静默错值 / Rejection path returns 0, no silent wrong value
        RETURN;                            // 快速失败出口，不再累加（Fast-fail exit, no further accumulation）
    END_IF

    uResult := uResult + USINT_TO_UINT(uDigit) * uWeight; // 位权累加：数值 × 当位权值（显式标准转换函数）/ Weighted accumulation with the standard explicit conversion
    uWeight := uWeight * DL_BCD_RADIX;     // 权值升位：1 → 10 → 100 → 1000 / Weight steps up: 1 -> 10 -> 100 -> 1000
END_FOR

(*------------------------------------------------------------------------------
 * 段 3｜结果回写（边界 B4）：纯函数出口唯一，无副作用
 *      Result write-back: single exit of the pure function, no side effect
 *      验收向量：16#0123 → 123；16#9999 → 9999；16#001A → 0 且置 0001_0105
 *      Acceptance vectors: 16#0123 -> 123; 16#9999 -> 9999; 16#001A -> 0 with 0001_0105
 *      上界自证：4 个半字节全 9 时 uResult = 9999 < 65535（UINT 域），无溢出
 *      Upper-bound proof: all-9 nibbles give 9999 < 65535 (UINT domain), no overflow
 *-----------------------------------------------------------------------------*)
FC_DL_BcdToWord := uResult;                // 全部半字节合法，返回累加结果 / All nibbles legal, return accumulated result
END_FUNCTION

(* ---- FC_DL_BinarySearchLReal.st ---- *)
(*==============================================================================
 * 组件名称 (Component)  : FC_DL_BinarySearchLReal
 * 所属子库 (Sublibrary) : DL_MathData
 * 当前版本 (Version)    : 1.0.1
 * 分类/来源标签         : lgf-datahandling（T2-1 LGF Data Handling 组回补）
 * 作者/日期             : Daoli Library / 2026-11-15
 * 兼容性   (Platform)   : CODESYS 3.5 / TwinCAT 3 / 汇川 InoProShop / Machine Expert
 *                         仅依赖 Standard.library（ABS），纯函数无状态
 * 功能简介 (Function)   : 对升序 LREAL 数组做经典二分查找，返回首个命中索引
 *                         （元素下标），未命中返回 -1；无状态、无副作用纯函数。
 *                         与 FB_DL_ArraySearchFirst 职责分离：
 *                         本块 = 升序数组 O(log n) 快速查找（要求调用方保证有序）；
 *                         线性块 = 无序数组 O(n) 通用查找。
 *                         典型现场用途：标定表按给定工程量反查断点槽位、
 *                         报警限值表按测量值定位档位区间、配方参数有序索引。
 * 开源溯源 (Origin)     : 原创实现（参考 LGF 公开手册 Data Handling 分类中
 *                         数组查找族的功能分类与参数域），只借分类/参数域/命名，
 *                         clean-room 实现，未复制任何源码。来源标签：lgf-datahandling。
 * 依赖     (Depends)    : 无 DL_ 内部依赖；Standard.library: ABS
 *
 * 【接口契约 / Interface contract】
 *   返回值：命中索引 [元素下标]，未命中 = -1。
 *   输入  ：afSorted 升序数组（调用方保证有序，VAR_IN_OUT 注入避免复制）；
 *           nCount 有效元素数；fTarget 目标值。
 *   输出  ：bFound 命中标志（与返回值同真相：TRUE 恒伴随返回值 >= 0）。
 *   纪律  ：纯函数同输入同输出；无内部状态；可安全放进 IF 表达式与
 *           多任务环境（无共享可变状态）。
 *
 * 【使用示例 / Usage example】
 *   VAR
 *       afCalTab : ARRAY[0..1023] OF LREAL;     // 升序标定表
 *       nSlot    : DINT;                        // 命中槽位
 *       bHit     : BOOL;                        // 命中标志
 *   END_VAR
 *   nSlot := FC_DL_BinarySearchLReal(afSorted := afCalTab,
 *                                    nCount := nRows, fTarget := fMeas,
 *                                    bFound => bHit);
 *   IF NOT bHit THEN
 *       nSlot := -1;    // 未命中走线性插值等后备逻辑
 *   END_IF
 *
 * 【选型对照 / Selection guide】
 *   本块（BinarySearchLReal）：升序数组、O(log n)、1024 元素最多 11 次比较、
 *                             不校验有序（契约责任在调用方）、无全量计数。
 *   FB_DL_ArraySearchFirst  ：无序可用、O(n) 单遍、支持全量计数与前缀搜索。
 *   高频轮询查找（每周期都查）选本块；低频事件查找 / 无序数据选线性块。
 *
 * 【算法与实时性披露 / Algorithm and timing disclosure】
 *   经典闭区间二分：每轮比较中点元素，命中即返；未命中按目标在左 / 右
 *   半区间收缩。DL_BS_MAX = 1024 时理论最大迭代 11 次（log2(1024) 向上取整），
 *   LREAL 比较约百纳秒级，单次调用总耗时微秒级以下，可放心放进每周期轮询。
 *   WHILE 循环配 64 次守护计数器（理论值的约 6 倍裕度），杜绝死循环。
 *
 * 验收向量 (Acceptance) : （afSorted = {1.5, 2.5, 3.5, 4.5, 5.5}，nCount = 5）
 *   V1 fTarget = 3.5 → 返回 2，bFound TRUE（中部命中）
 *   V2 fTarget = 1.5 → 返回 0，bFound TRUE（下边界命中）
 *   V3 fTarget = 5.5 → 返回 4，bFound TRUE（上边界命中）
 *   V4 fTarget = 3.6 → 返回 -1，bFound FALSE（带内未命中，容差外）
 *   V5 fTarget = 0.5 → 返回 -1，bFound FALSE（低于全域）
 *
 * 【V1 逐轮迭代推演 / Iteration trace of V1】
 *   轮次 ｜ nLo ｜ nHi ｜ nMid ｜ 探测值 ｜ 判定
 *   1    ｜ 0   ｜ 4    ｜ 2     ｜ 3.5    ｜ 容差命中 → 返回 2（1 轮即中）
 * 【V4 逐轮迭代推演 / Iteration trace of V4】（fTarget = 3.6）
 *   轮次 ｜ nLo ｜ nHi ｜ nMid ｜ 探测值 ｜ 判定
 *   1    ｜ 0   ｜ 4    ｜ 2     ｜ 3.5    ｜ 3.5 < 3.6 → 收缩右半 nLo=3
 *   2    ｜ 3   ｜ 4    ｜ 3     ｜ 4.5    ｜ 4.5 > 3.6 → 收缩左半 nHi=2
 *   3    ｜ nLo=3 > nHi=2 → 区间塌缩，WHILE 退出，返回 -1（3 轮收敛）
 *
 * 【重复值语义声明 / Duplicate-value semantics】
 *   数组含重复目标值时返回其中任一命中下标（经典二分不保证首个），
 *   需要"首个命中"语义的场合请改用 FB_DL_ArraySearchFirst（线性块），
 *   该契约与线性块的"首个命中"形成互补，选型时按语义需求取舍。
 *
 * 【常见误用清单 / Common misuse checklist】
 *   M1 对无序数组调用 → 返回值无意义（B1 契约责任），先排序再查；
 *   M2 nCount 传数组全长而实际只装了前 n 行 → 残留旧数据可能误命中，
 *      按实际装载行数传参；
 *   M3 把返回值直接当下标写数组而不查 bFound → 未命中时 -1 会被当
 *      "最后一个元素"（部分平台负下标越界），必须先判 bFound；
 *   M4 用本块结果做浮点精确相等断言 → 命中本身已是容差口径，
 *      后续再判等请沿用同一容差常量，勿混用严格判等；
 *   M5 在扫描周期内对同一表反复排序+查找 → 排序成本远高于查找本身，
 *      排序一次后缓存"已有序"标志再高频查找。
 * 故障码表 (Error codes):
 *   16#0001_010F  nCount 越界，已钳位到 0..DL_BS_MAX（信息级，查找照常执行）
 *   16#0001_0206  二分守护计数超限或下标兜底触发，强制返回未命中
 *                 （故障级，理论不可达）
 *                 【码位终审】原拟 0002_0101 / 0002_0201 与 DL_Algo PID 族
 *                 （FB_DL_PidController 0002_0101 输出饱和、FB_DL_CascadePid
 *                 0002_0201 副设定钳位）冲突，且 0002_01xx 段已由 DL_Algo
 *                 PID 族登记；DL_MathData 依公约 0.7 归 0001_xxxx 段，
 *                 R9 终审顺延至 0001_010F / 0001_0206（与既有 0101~010F、
 *                 0201~0212 逐条比对无冲突）。
 * 红线自检 (Redline)    : R1 ✓ 零全局存储 / 零外部变量引用 ｜ R2 ✓ 零物理地址直写
 *                         R3 ✓ 纯 IEC 61131-3 ｜ R4 ✓ nCount 钳位 + 中点防溢出 + 守护计数 + 容差判等 + 空表直退
 *                         R5 ✓ 全变量中英双语同行注释 ｜ R6 ✓ 纯函数无状态（R6 状态机 N/A）
 *                         R7 ✓ 无定时器 / 边沿实例（R7 N/A）
 * 边界契约 (Boundaries):
 *   B1 调用方保证数组升序有序，本函数不校验全序（校验需 O(n)，会摧毁 O(log n) 价值）；
 *      无序输入的返回值无意义，属调用方契约责任，头注释写死。
 *   B2 中点计算固定写法 nMid := nLo + (nHi - nLo) / 2，防 (nLo + nHi) 溢出，
 *      DINT 域内安全——二分实现中最常见的溢出缺陷，此处从写法上根除。
 *   B3 守护上限 64 次：DL_BS_MAX = 1024 理论最大迭代 11 次，64 为约 6 倍裕度，
 *      超限视为平台异常强制退出，bFound FALSE 返回 -1，绝不死循环。
 *   B4 命中判据 ABS(afSorted[nMid] - fTarget) < DL_FLOAT_EPS，禁浮点直接判等；
 *      区间收缩判据用严格大于 / 小于，与容差判等正交不冲突。
 *   B5 nCount = 0（空表）直接返回 -1，合法工况不置故障码。
 * 修订历史 (Revision)   :
 *   2026-11-15  v1.0.0  首版落盘（Round 09 · 泳道 A · Level 0 原子族回补）
 *   2026-11-15  v1.0.1  终审修复：补声明缺失的 uErrorId 输出引脚（原 1.0.0 在
 *                       函数体内五处读写 uErrorId 却未声明，三平台均编译失败）；
 *                       故障码 0002_0101/0002_0201 与 DL_Algo PID 族冲突，
 *                       顺延至 0001_010F / 0001_0206（同段位归口 DL_MathData）
 *============================================================================*)
FUNCTION FC_DL_BinarySearchLReal : DINT    // 返回命中索引 [元素下标]，未命中 = -1 / Hit index, -1 when not found
VAR_IN_OUT
    afSorted   : ARRAY[0..DL_BS_MAX-1] OF LREAL;  // 升序数组（调用方保证有序，本函数不校验全序）/ Ascending array, sorted by the caller
END_VAR
VAR_INPUT
    nCount     : DINT;                 // 有效元素数 [个]，0..DL_BS_MAX，越界钳位 / Valid element count [items], clamped
    fTarget    : LREAL;                // 目标值 [工程单位随应用] / Target value [EU by application]
END_VAR
VAR_OUTPUT
    bFound     : BOOL;                 // 命中标志，与返回值同真相源 / Hit flag, same truth as the return value
    uErrorId   : UDINT;                // 故障码，0 = 无故障（0001_010F 钳位信息级 / 0001_0206 守护故障级）/ Error code, 0 = no error
END_VAR
VAR
    nLo        : DINT;                 // 区间下界索引（闭区间）/ Interval lower bound index, inclusive
    nHi        : DINT;                 // 区间上界索引（闭区间）/ Interval upper bound index, inclusive
    nMid       : DINT;                 // 中点索引 / Midpoint index
    nGuard     : DINT;                 // 循环防死锁守护计数器 [次] / Loop guard counter [iterations]
    nCountEff  : DINT;                 // 钳位后的有效元素数 [个] / Effective clamped element count [items]
    fProbe     : LREAL;                // 当前探测点元素值缓存 / Probed element value cache
END_VAR
VAR CONSTANT
    DL_BS_MAX   : DINT := 1024;        // 数组容量上限 [元素]，必须与数组维度一致 / Array capacity limit, must match the dimension
    DL_BS_GUARD : DINT := 64;          // 二分守护上限 [次]，理论 11 次 × 约 6 倍裕度 / Binary guard limit, ~6x margin of theory
    DL_FLOAT_EPS: LREAL := 1.0E-9;     // LREAL 判等容差，禁浮点直接判等 / LREAL equality tolerance
END_VAR

(*------------------------------------------------------------------------------
 * 段 1｜缺省返回：未命中语义（-1 / FALSE），故障码清零
 *      Default return: miss semantics, error code cleared
 *      缺省即失败语义：任何提前退出路径都自动携带"未命中"，不会误报成功
 *-----------------------------------------------------------------------------*)
FC_DL_BinarySearchLReal := -1;
bFound    := FALSE;
uErrorId  := 16#0000_0000;

(*------------------------------------------------------------------------------
 * 段 2｜范围钳位与空表直退（边界 B5）：nCount = 0 合法直退不置故障
 *      Range clamp and empty-table early exit
 *-----------------------------------------------------------------------------*)
IF (nCount < 0) OR (nCount > DL_BS_MAX) THEN
    IF nCount < 0 THEN
        nCountEff := 0;         // 负数视作空表 / Negative treated as empty
    ELSE
        nCountEff := DL_BS_MAX; // 超上限截断 / Overflow truncated
    END_IF
    uErrorId := 16#0001_010F;   // 信息级：范围越界已钳位 / Info: range clamped
ELSE
    nCountEff := nCount;        // 合法范围直通 / Legal range passes through
END_IF

IF nCountEff <= 0 THEN
    RETURN;                     // 空表：合法工况，保持缺省未命中返回
END_IF

(*------------------------------------------------------------------------------
 * 段 3｜经典二分主体（边界 B2/B3/B4）：闭区间 [nLo, nHi]，中点防溢出写法，
 *      守护计数超限强制退出，命中判据用容差
 *      Classic binary search on a closed interval with overflow-safe midpoint
 *-----------------------------------------------------------------------------*)
nLo    := 0;                    // 闭区间下界从 0 起 / Closed lower bound from 0
nHi    := nCountEff - 1;        // 闭区间上界到末元素 / Closed upper bound at the last element
nGuard := 0;                    // 守护计数清零 / Guard counter cleared

WHILE (nLo <= nHi) AND (nGuard < DL_BS_GUARD) DO
    nGuard := nGuard + 1;       // 每轮累加，超限即退出（B3）

    (* 中点防溢出固定写法：不写 (nLo + nHi) / 2，DINT 极值下不回绕（B2） *)
    nMid := nLo + (nHi - nLo) / 2;

    (* 下标先判界再访问（红线 R4）：区间不变式已保证，仍显式兜底 *)
    IF (nMid >= 0) AND (nMid < DL_BS_MAX) THEN
        fProbe := afSorted[nMid];   // 取中点元素 / Probe the midpoint element
    ELSE
        uErrorId := 16#0001_0206;   // 故障级：下标越界兜底 / Fault: index guard tripped
        RETURN;
    END_IF

    IF ABS(fProbe - fTarget) < DL_FLOAT_EPS THEN
        FC_DL_BinarySearchLReal := nMid;    // 命中：返回当前下标 / Hit: return the index
        bFound := TRUE;
        RETURN;
    ELSIF fProbe < fTarget THEN
        nLo := nMid + 1;            // 目标在右半区间 / Target in the right half
    ELSE
        nHi := nMid - 1;            // 目标在左半区间 / Target in the left half
    END_IF
END_WHILE

(*------------------------------------------------------------------------------
 * 段 4｜守护超限兜底（边界 B3）：理论不可达，置故障级码保持未命中返回
 *      Guard-exceeded fallback: theoretically unreachable, fault code kept
 *-----------------------------------------------------------------------------*)
IF nGuard >= DL_BS_GUARD THEN
    uErrorId := 16#0001_0206;   // 故障级：守护超限 / Fault: guard exceeded
END_IF
END_FUNCTION
